// ---- TEST/LOGGING/PROCESSOR/UTILS/FB_LogRecordProcessor_ForBatchInspection.TcPOU
(*
	Processor test double that exposes the batch processor's record queue for assertions.
	Unlike FB_LogRecordProcessor_ForRecordsInspection it does NOT override
	onEmit, so tests exercise the real batch grouping behavior.
*)
FUNCTION_BLOCK FB_LogRecordProcessor_ForBatchInspection EXTENDS FB_LogRecordProcessor_Batch

// explicitly run the batch processor body so tests exercise the flush logic
SUPER^();

PROPERTY records : REFERENCE TO FB_LogRecordQueue
GET
records REF= THIS^._records;
END_GET
END_PROPERTY

END_FUNCTION_BLOCK

// ---- TEST/LOGGING/EXPORTING/FB_TestLogExporters.TcPOU
(* Tests the contract between a caller's batch and a log exporter. *)
FUNCTION_BLOCK FB_TestLogExporters EXTENDS FB_TestSuite

THIS^.testExportSerializesWholeBatch();

(*
	export takes ownership of every record in the caller's batch and passes them to the serializer, so the
	caller holds nothing the exporter will release. Grouping by resource and scope is tested in FB_TestProtoJsonSerializer.
*)
METHOD testExportSerializesWholeBatch : REFERENCE TO FB_Test
VAR CONSTANT
	RECORD_COUNT: UDINT := 2;  // more than one, so the whole batch has to move, not just its head
END_VAR
VAR
	resource: FB_Resource(schemaUrl:='');
	provider: FB_LoggerProvider(resource:=resource);
	scope: FB_InstrumentationScope(name:='exporter.test', version:='1.0.0', schemaUrl:='');
	logger: FB_Logger(scope:=scope, provider:=provider);
	processor: FB_LogRecordProcessor_ForRecordsInspection(
		maxQueueSize:=0,
		scheduledDelayMillis:=1000,
		maxExportBatchSize:=512,
		exporter:=0
	);
	exporter: FB_LogRecordExporter_File_ForSerializationInspection;
	serialized: REFERENCE TO FB_LogRecordProtoJsonSerializer;
	emitSucceeded: BOOL;
	emitFailureReason: E_LoggerFailureReason;
	exporterFailureReason: E_LogRecordExporterFailureReason;
	exportSucceeded: BOOL;
	resourceLogs: SJsonValue;
	_idx: UDINT;
END_VAR
TcUnit.TEST('testExportSerializesWholeBatch');
	// arrange: the processor collects a batch emitted through the logger; its resource and scope do not matter here
	processor.free();
	FOR _idx := 1 TO RECORD_COUNT DO
		emitSucceeded := logger
			.startLogRecord(severityNumber:=E_SeverityNumber.INFO)
			.setTimestamp(TO_ULINT(_idx))
			.emit(failureResult=>emitFailureReason);
		THIS^.AssertTrue(emitSucceeded, 'Expected the logger to emit the record');
	END_FOR
	provider
		.stageProcessor(processor)
		.tick();
	THIS^.AssertEquals_UDINT(RECORD_COUNT, processor.records.count, 'Expected the processor to collect every emitted record');

	// act
	exportSucceeded := processor.exportRecords(exporter:=exporter, failureReason=>exporterFailureReason);

	// assert: the exporter owns the whole batch and serialized it
	THIS^.AssertTrue(
		exportSucceeded
		AND_THEN processor.records.count = 0
		AND_THEN exporterFailureReason = E_LogRecordExporterFailureReason.NA,
		'Expected export to succeed with no failure reason and take every record out of the batch'
	);
	serialized REF= exporter.serializer;
	resourceLogs := serialized.parser.FindMember(serialized.jsonValue, 'resourceLogs');
	THIS^.AssertTrue(resourceLogs <> 0 AND_THEN serialized.parser.IsArray(resourceLogs), 'Expected the exporter to serialize the batch into a resourceLogs array');

	exporter.free();
	processor.free();
TcUnit.TEST_FINISHED();
END_METHOD

END_FUNCTION_BLOCK

// ---- TEST/LOGGING/PROCESSOR/UTILS/FB_LogRecordProcessor_ForRecordsInspection.TcPOU
(* Processor test double that retains emitted records for assertions. *)
// lastOperationSucceeded and failureResult are inherited from FB_LogRecordProcessor_Batch
FUNCTION_BLOCK FB_LogRecordProcessor_ForRecordsInspection EXTENDS FB_LogRecordProcessor_Batch

METHOD exportRecords : BOOL
VAR_INPUT
	exporter: REFERENCE TO FB_LogRecordExporter_Base;
END_VAR
VAR_OUTPUT
	failureReason: E_LogRecordExporterFailureReason;
END_VAR
exportRecords := exporter.export(
	logRecords:=THIS^._records,
	count:=THIS^._records.count,
	failureReason=>failureReason
);
END_METHOD

(*
	Retains every emitted record for assertions, whether or not an exporter is
	bound. FB_LogRecordProcessor_Batch.onEmit deliberately skips the clone and
	the queue push when it has no exporter; this double overrides that so a test
	can collect records and hand them to an exporter itself via exportRecords.
*)
METHOD onEmit
VAR_INPUT
	logRecord: REFERENCE TO FB_LogRecord;
END_VAR
VAR
	_pRecord: POINTER TO FB_LogRecord;
	_cloneFailureResult: E_LogRecordCloneFailureReason;
	_queueFailureReason: E_LogRecordQueueFailureReason;
END_VAR
THIS^.enrich(logRecord);

_pRecord := 0;
IF NOT logRecord.cloneTo(pDest:=_pRecord, failureReason=>_cloneFailureResult) THEN
	IF _pRecord <> 0 THEN _pRecord^.delete(pSelf:=_pRecord); END_IF
	THIS^.lastOperationSucceeded := FALSE;
	THIS^.failureResult := E_LogRecordProcessorFailureReason.RECORD_CLONE_FAILURE;
	RETURN;
END_IF

IF NOT THIS^._records.push(pValue:=_pRecord, failureReason=>_queueFailureReason) THEN
	_pRecord^.delete(pSelf:=_pRecord);
	THIS^.lastOperationSucceeded := FALSE;
	THIS^.failureResult := E_LogRecordProcessorFailureReason.QUEUE_PUSH_FAILURE;
	RETURN;
END_IF

THIS^.lastOperationSucceeded := TRUE;
THIS^.failureResult := E_LogRecordProcessorFailureReason.NA;
END_METHOD

PROPERTY records : REFERENCE TO FB_LogRecordQueue
GET
records REF= THIS^._records;
END_GET
END_PROPERTY

END_FUNCTION_BLOCK

// ---- TEST/LOGGING/EXPORTING/UTILS/FB_LogRecordExporter_File_ForSerializationInspection.TcPOU
(* Exporter test double that serializes accepted records without destination I/O. *)
FUNCTION_BLOCK FB_LogRecordExporter_File_ForSerializationInspection EXTENDS FB_LogRecordExporter_Base
VAR_OUTPUT
	serializer: FB_LogRecordProtoJsonSerializer;
END_VAR
VAR
	_serializationFailureReason: E_ProtoJsonSerializerFailureReason;
END_VAR

METHOD export : BOOL
VAR_IN_OUT
	logRecords: FB_LogRecordQueue;
END_VAR
VAR_INPUT
	count: UDINT;
END_VAR
VAR_OUTPUT
	failureReason: E_LogRecordExporterFailureReason;
END_VAR
_serializationFailureReason := E_ProtoJsonSerializerFailureReason.NA;
export := SUPER^.export(
	logRecords:=logRecords,
	count:=count,
	failureReason=>failureReason
);
IF NOT export THEN
	RETURN;
END_IF

IF NOT THIS^.serializer.serializeLogsData(
	logRecords:=THIS^._records,
	failureReason=>_serializationFailureReason
) THEN
	failureReason := E_LogRecordExporterFailureReason.SERIALIZATION_FAILURE;
	export := FALSE;
END_IF
THIS^.free();
END_METHOD

METHOD isBusy : BOOL
isBusy := FALSE;
END_METHOD

METHOD tick : BOOL
VAR_OUTPUT
	failureReason: E_LogRecordExporterFailureReason;
END_VAR
failureReason := E_LogRecordExporterFailureReason.NA;
tick := TRUE;
END_METHOD

END_FUNCTION_BLOCK

// ---- TEST/LOGGING/LOG_RECORD/FB_TestLogRecord.TcPOU
(* Tests log record ownership and cloning. *)
FUNCTION_BLOCK FB_TestLogRecord EXTENDS FB_TestSuite
VAR_INPUT
END_VAR
VAR_OUTPUT
END_VAR
VAR
END_VAR

THIS^.testCloneToIsIndependent();

(* cloneTo deep copies a record, its resource, scope and every owned value, so a processor can keep the clone after the logger frees the source. Cloning into an assigned destination is refused so the existing record is not leaked. *)
METHOD testCloneToIsIndependent : REFERENCE TO FB_Test
VAR_INPUT
END_VAR
VAR
	resource: FB_Resource('resource.schema');
	provider: FB_LoggerProvider(resource);
	scope: FB_InstrumentationScope('scope.name', '1.0.0', 'scope.schema');
	logger: FB_Logger(scope, provider);
	timestamp: ULINT := 123456789;
	traceIdBytes: ARRAY [0..15] OF BYTE := [0, 1, 2, 3, 4, 5, 6, 7, 8, 9, 10, 11, 12, 13, 14, 15];
	spanIdBytes: ARRAY [0..7] OF BYTE := [16, 17, 18, 19, 20, 21, 22, 23];
	cloneSuccess: BOOL;
	cloneFailureResult: E_LogRecordCloneFailureReason;
	attributesSuccess: BOOL;
	attributesFailureReason: E_AttributesFailureReason;
	pClone: POINTER TO FB_LogRecord;
	pSourceResourceAttribute: POINTER TO FB_KeyValue;
	pClonedResourceAttribute: POINTER TO FB_KeyValue;
	pSourceScopeAttribute: POINTER TO FB_KeyValue;
	pClonedScopeAttribute: POINTER TO FB_KeyValue;
	pSourceRecordAttribute: POINTER TO FB_KeyValue;
	pClonedRecordAttribute: POINTER TO FB_KeyValue;
	pSourceString: POINTER TO FB_String;
	pClonedString: POINTER TO FB_String;
END_VAR
TcUnit.TEST('testCloneToIsIndependent');
	// Arrange: a source record with event name, body, IDs and one attribute at each level
	attributesSuccess := resource.attributes.setStringAttribute(
		key:='resource.key',
		value:='resource.value',
		failureReason=>attributesFailureReason
	);
	THIS^.AssertTrue(attributesSuccess, 'Expected resource attribute creation to succeed');
	attributesSuccess := scope.attributes.setStringAttribute(
		key:='scope.key',
		value:='scope.value',
		failureReason=>attributesFailureReason
	);
	THIS^.AssertTrue(attributesSuccess, 'Expected scope attribute creation to succeed');

	logger
		.startLogRecord(severityNumber:=E_SeverityNumber.INFO)
		.setTimestamp(timestamp)
		.setEventName('record.event')
		.setBody('record.body')
		._setTraceId(ADR(traceIdBytes), SIZEOF(traceIdBytes))
		._setSpanId(ADR(spanIdBytes), SIZEOF(spanIdBytes))
		._setFlags(16#01)  // sampled
		.setStringAttribute('record.key', 'record.value');
	THIS^.AssertTrue(logger.pLogRecord <> 0, 'Expected startLogRecord to build a source log record');

	// Clone: the first clone succeeds, a second into the same destination is refused
	IF logger.pLogRecord <> 0 THEN
		// no builder sets droppedAttributesCount; set by hand so the clone has a non-default value to copy
		logger.pLogRecord^.droppedAttributesCount := 4;
		cloneSuccess := logger.pLogRecord^.cloneTo(
			pDest:=pClone,
			failureReason=>cloneFailureResult
		);
		THIS^.AssertTrue(cloneSuccess, 'Expected log record clone to succeed');
		THIS^.AssertTrue(pClone <> 0, 'Expected a cloned log record');
		THIS^.AssertTrue(pClone <> logger.pLogRecord, 'Expected a distinct log record allocation');

		cloneSuccess := logger.pLogRecord^.cloneTo(
			pDest:=pClone,
			failureReason=>cloneFailureResult
		);
		THIS^.AssertFalse(cloneSuccess, 'Expected cloning into an assigned destination to fail');
		THIS^.AssertTrue(
			cloneFailureResult = E_LogRecordCloneFailureReason.DESTINATION_ALREADY_ASSIGNED,
			'Expected the DESTINATION_ALREADY_ASSIGNED reason when cloning into an assigned destination'
		);
	END_IF

	// Copied fields: equal values, distinct allocations for every owned value
	IF pClone <> 0 AND_THEN logger.pLogRecord <> 0 THEN
		THIS^.AssertTrue(pClone^.severityNumber = logger.pLogRecord^.severityNumber, 'Expected severity number to be cloned');
		THIS^.AssertTrue(pClone^.timestamp = logger.pLogRecord^.timestamp, 'Expected timestamp to be cloned');
		THIS^.AssertEquals_UDINT(logger.pLogRecord^.droppedAttributesCount, pClone^.droppedAttributesCount, 'Expected dropped record attribute count to be cloned');
		THIS^.AssertEquals_STRING(logger.pLogRecord^.resource.schemaUrl, pClone^.resource.schemaUrl, 'Expected resource schema URL to be cloned');
		THIS^.AssertEquals_UDINT(logger.pLogRecord^.resource.droppedAttributesCount, pClone^.resource.droppedAttributesCount, 'Expected dropped resource attribute count to be cloned');
		THIS^.AssertEquals_STRING(logger.pLogRecord^.scope.name, pClone^.scope.name, 'Expected scope name to be cloned');
		THIS^.AssertEquals_STRING(logger.pLogRecord^.scope.version, pClone^.scope.version, 'Expected scope version to be cloned');
		THIS^.AssertEquals_STRING(logger.pLogRecord^.scope.schemaUrl, pClone^.scope.schemaUrl, 'Expected scope schema URL to be cloned');
		THIS^.AssertEquals_UDINT(logger.pLogRecord^.scope.droppedAttributesCount, pClone^.scope.droppedAttributesCount, 'Expected dropped scope attribute count to be cloned');
		THIS^.AssertTrue(pClone^.eventName <> logger.pLogRecord^.eventName, 'Expected event name allocation to be cloned');
		THIS^.AssertTrue(pClone^.eventName^.pString <> logger.pLogRecord^.eventName^.pString, 'Expected event name string allocation to be cloned');
		THIS^.AssertEquals_STRING(logger.pLogRecord^.eventName^.pString^, pClone^.eventName^.pString^, 'Expected event name value to be cloned');
		THIS^.AssertTrue(pClone^.traceId <> logger.pLogRecord^.traceId, 'Expected trace ID allocation to be cloned');
		THIS^.AssertTrue(MEMCMP(ADR(pClone^.traceId^.bytes), ADR(logger.pLogRecord^.traceId^.bytes), SIZEOF(pClone^.traceId^.bytes)) = 0, 'Expected trace ID value to be cloned');
		THIS^.AssertEquals_UDINT(1, pClone^.flags, 'Expected the sampled trace flag to be cloned');
		THIS^.AssertTrue(pClone^.spanId <> logger.pLogRecord^.spanId, 'Expected span ID allocation to be cloned');
		THIS^.AssertTrue(MEMCMP(ADR(pClone^.spanId^.bytes), ADR(logger.pLogRecord^.spanId^.bytes), SIZEOF(pClone^.spanId^.bytes)) = 0, 'Expected span ID value to be cloned');
		THIS^.AssertTrue(pClone^.body <> logger.pLogRecord^.body, 'Expected body allocation to be cloned');
		pSourceString := logger.pLogRecord^.body;
		pClonedString := pClone^.body;
		THIS^.AssertTrue(pClonedString^.pString <> pSourceString^.pString, 'Expected body string allocation to be cloned');
		THIS^.AssertEquals_STRING(pSourceString^.pString^, pClonedString^.pString^, 'Expected body value to be cloned');

		// Attributes: each level's attribute, key and value are new allocations
		logger.pLogRecord^.resource.attributes.reset();
		pClone^.resource.attributes.reset();
		pSourceResourceAttribute := logger.pLogRecord^.resource.attributes.next();
		pClonedResourceAttribute := pClone^.resource.attributes.next();
		THIS^.AssertTrue(pSourceResourceAttribute <> 0, 'Expected the source record to have a resource attribute');
		THIS^.AssertTrue(pClonedResourceAttribute <> 0, 'Expected the cloned record to have a resource attribute');
		IF pSourceResourceAttribute <> 0 AND_THEN pClonedResourceAttribute <> 0 THEN
			THIS^.AssertTrue(pClonedResourceAttribute <> pSourceResourceAttribute, 'Expected resource attribute allocation to be cloned');
			THIS^.AssertTrue(pClonedResourceAttribute^.pKey <> pSourceResourceAttribute^.pKey, 'Expected resource attribute key allocation to be cloned');
			THIS^.AssertTrue(pClonedResourceAttribute^.pVal <> pSourceResourceAttribute^.pVal, 'Expected resource attribute value allocation to be cloned');
		END_IF

		logger.pLogRecord^.scope.attributes.reset();
		pClone^.scope.attributes.reset();
		pSourceScopeAttribute := logger.pLogRecord^.scope.attributes.next();
		pClonedScopeAttribute := pClone^.scope.attributes.next();
		THIS^.AssertTrue(pSourceScopeAttribute <> 0, 'Expected the source record to have a scope attribute');
		THIS^.AssertTrue(pClonedScopeAttribute <> 0, 'Expected the cloned record to have a scope attribute');
		IF pSourceScopeAttribute <> 0 AND_THEN pClonedScopeAttribute <> 0 THEN
			THIS^.AssertTrue(pClonedScopeAttribute <> pSourceScopeAttribute, 'Expected scope attribute allocation to be cloned');
			THIS^.AssertTrue(pClonedScopeAttribute^.pKey <> pSourceScopeAttribute^.pKey, 'Expected scope attribute key allocation to be cloned');
			THIS^.AssertTrue(pClonedScopeAttribute^.pVal <> pSourceScopeAttribute^.pVal, 'Expected scope attribute value allocation to be cloned');
		END_IF

		logger.pLogRecord^.attributes.reset();
		pClone^.attributes.reset();
		pSourceRecordAttribute := logger.pLogRecord^.attributes.next();
		pClonedRecordAttribute := pClone^.attributes.next();
		THIS^.AssertTrue(pSourceRecordAttribute <> 0, 'Expected the source record to have a record attribute');
		THIS^.AssertTrue(pClonedRecordAttribute <> 0, 'Expected the cloned record to have a record attribute');
		IF pSourceRecordAttribute <> 0 AND_THEN pClonedRecordAttribute <> 0 THEN
			THIS^.AssertTrue(pClonedRecordAttribute <> pSourceRecordAttribute, 'Expected record attribute allocation to be cloned');
			THIS^.AssertTrue(pClonedRecordAttribute^.pKey <> pSourceRecordAttribute^.pKey, 'Expected record attribute key allocation to be cloned');
			THIS^.AssertTrue(pClonedRecordAttribute^.pVal <> pSourceRecordAttribute^.pVal, 'Expected record attribute value allocation to be cloned');
		END_IF
	END_IF

	// Independence: the clone keeps its values after the logger frees the source
	logger.free();
	THIS^.AssertTrue(logger.pLogRecord = 0, 'Expected source log record to be deleted');

	IF pClone <> 0 THEN
		THIS^.AssertEquals_STRING('record.event', pClone^.eventName^.pString^, 'Expected cloned event name to survive source deletion');
		pClonedString := pClone^.body;
		THIS^.AssertEquals_STRING('record.body', pClonedString^.pString^, 'Expected cloned body to survive source deletion');
		THIS^.AssertEquals_UDINT(1, pClone^.resource.attributes.count, 'Expected cloned resource attributes to survive source deletion');
		THIS^.AssertEquals_UDINT(1, pClone^.scope.attributes.count, 'Expected cloned scope attributes to survive source deletion');
		THIS^.AssertEquals_UDINT(1, pClone^.attributes.count, 'Expected cloned record attributes to survive source deletion');
		pClone^.delete(pSelf:=pClone);
	END_IF
TcUnit.TEST_FINISHED();
END_METHOD

END_FUNCTION_BLOCK

// ---- TEST/LOGGING/SERIALIZATION/FB_TestProtoJsonSerializer.TcPOU
(* Tests that the base and log-record ProtoJSON serializers write the OTLP/JSON wire form: field encodings, failure reasons, and resource/scope grouping. *)
FUNCTION_BLOCK FB_TestProtoJsonSerializer EXTENDS FB_TestSuite

THIS^.testSerializeNumberValues();
THIS^.testSerializeLogRecord();
THIS^.testSerializeLogRecordWithoutTraceIdOmitsFlags();
THIS^.testSerializeRejectsNullInputs();
THIS^.testSerializeLogsDataGroupsByResourceAndScope();

(* A null log-record pointer or a null member key fails serialization with its own failure reason,
   so a caller can tell a missing record from a serializer misuse instead of writing broken JSON. *)
METHOD testSerializeRejectsNullInputs : REFERENCE TO FB_Test
VAR
	serializer: FB_LogRecordProtoJsonSerializer;
	root: SJsonValue;
	records: SJsonValue;
	pRecord: POINTER TO FB_LogRecord;
	serializationSucceeded: BOOL;
	failureReason: E_ProtoJsonSerializerFailureReason;
END_VAR
TcUnit.TEST('testSerializeRejectsNullInputs');
	root := serializer.parser.NewDocument();
	root := serializer.parser.SetObject(root);
	records := serializer.parser.AddArrayMember(root, 'logRecords', 0);

	// pRecord is deliberately left 0.
	serializationSucceeded := serializer.serializeLogRecord(
		v:=records,
		pLogRecord:=pRecord,
		failureReason=>failureReason
	);
	THIS^.AssertFalse(serializationSucceeded, 'Expected a null log-record pointer to fail serialization');
	THIS^.AssertTrue(
		failureReason = E_ProtoJsonSerializerFailureReason.LOG_RECORD_POINTER_NULL,
		'Expected LOG_RECORD_POINTER_NULL as the failure reason for a null log record'
	);

	// pKey is deliberately 0.
	serializationSucceeded := serializer.serializeUint32Value(
		v:=root,
		pKey:=0,
		val:=1,
		failureReason=>failureReason
	);
	THIS^.AssertFalse(serializationSucceeded, 'Expected a null JSON member key to fail serialization');
	THIS^.AssertTrue(
		failureReason = E_ProtoJsonSerializerFailureReason.KEY_POINTER_NULL,
		'Expected KEY_POINTER_NULL as the failure reason for a null member key'
	);
TcUnit.TEST_FINISHED();
END_METHOD

(* A record built through the logger serializes every field in its OTLP/JSON form: enums and fixed32 as numbers,
   64-bit integers as decimal strings, trace and span IDs as hex, and values as typed AnyValue objects. *)
METHOD testSerializeLogRecord : REFERENCE TO FB_Test
VAR
	resource: FB_Resource(schemaUrl:='');
	provider: FB_LoggerProvider(resource:=resource);
	scope: FB_InstrumentationScope(name:='motor1', version:='0.0.1a', schemaUrl:='');
	logger: FB_Logger(scope:=scope, provider:=provider);
	processor: FB_LogRecordProcessor_ForRecordInspection(0);
	serializer: FB_LogRecordProtoJsonSerializer();
	emitSuccess: BOOL;
	emitFailureResult: E_LoggerFailureReason;
	timestamp: ULINT := 1581452773000000789;
	traceId: ARRAY [0..15] OF BYTE := [0, 1, 2, 3, 4, 5, 6, 7, 8, 9, 10, 11, 12, 13, 14, 15];
	spanId: ARRAY [0..7] OF BYTE := [16, 17, 18, 19, 20, 21, 22, 23];
	durationMs: DINT := 42;
	temperature: LREAL := 21.5;
	pRecord: POINTER TO FB_LogRecord;
	root: SJsonValue;
	records: SJsonValue;
	obj: SJsonValue;
	member: SJsonValue;
	attributes: SJsonValue;
	attribute: SJsonValue;
	value: SJsonValue;
	actualString: STRING;
	serializationSucceeded: BOOL;
	serializerFailureReason: E_ProtoJsonSerializerFailureReason;
END_VAR
TcUnit.TEST('testSerializeLogRecord');
	processor.free();
	logger.free();

	// Create a representative record through the public logger API.
	logger
		.startLogRecord(severityNumber:=E_SeverityNumber.DEBUG)
		.setTimestamp(timestamp)
		.setEventName('Serialization Event')
		.setBody('This is a body string value')
		._setTraceId(ADR(traceId), SIZEOF(traceId))
		._setSpanId(ADR(spanId), SIZEOF(spanId))
		._setFlags(16#01)  // sampled
		.setStringAttribute('stats.label', 'pVal')
		.setNumberAttribute('stats.duration_ms', durationMs)
		.setNumberAttribute('stats.temperature', temperature);
	THIS^.AssertTrue(logger.pLogRecord <> 0, 'Expected the logger to hold a log record before emission');
	IF logger.pLogRecord <> 0 THEN
		// no builder sets droppedAttributesCount; set by hand to check it is written
		logger.pLogRecord^.droppedAttributesCount := 2;
	END_IF

	emitSuccess := logger.emit(failureResult=>emitFailureResult);
	THIS^.AssertTrue(emitSuccess, 'Expected log record emission to succeed');
	provider
		.stageProcessor(processor)
		.tick();
	THIS^.AssertTrue(processor.lastOperationSucceeded, 'Expected the inspection processor to capture the emitted record');
	THIS^.AssertTrue(logger.pLogRecord = 0, 'Expected emit to release the logger-owned record');
	pRecord := processor.pop();
	THIS^.AssertTrue(pRecord <> 0, 'Expected the processor to return the emitted record');
	IF pRecord <> 0 THEN

	// serializeLogRecord appends one LogRecord object to the supplied JSON array.
	root := serializer.parser.NewDocument();
	serializer.parser.SetObject(root);
	records := serializer.parser.AddArrayMember(root, 'logRecords', 0);
	serializationSucceeded := serializer.serializeLogRecord(
		v:=records,
		pLogRecord:=pRecord,
		failureReason=>serializerFailureReason
	);
	THIS^.AssertTrue(
		serializationSucceeded AND_THEN serializerFailureReason = E_ProtoJsonSerializerFailureReason.NA,
		'Expected LogRecord serialization to succeed without a failure reason'
	);
	obj := serializer.parser.GetArrayValueByIdx(records, 0);
		THIS^.AssertTrue(serializer.parser.IsObject(obj), 'Expected the logRecords array to hold one LogRecord object');

		// OTLP/JSON encodes enums and fixed32 values as numbers.
		// 5 is DEBUG; flags 1 is the sampled trace flag of the record's span.
		member := serializer.parser.FindMember(obj, 'severityNumber');
		THIS^.AssertEquals_UDINT(5, serializer.parser.GetUint(member), 'Expected severityNumber 5 (DEBUG) as a JSON number');
		actualString := serializer.parser.GetString(serializer.parser.FindMember(obj, 'severityText'));
		THIS^.AssertEquals_STRING('DEBUG', actualString, 'Expected severityText to be the severity enum name');
		THIS^.AssertEquals_UDINT(1, serializer.parser.GetUint(serializer.parser.FindMember(obj, 'flags')), 'Expected flags 1 (sampled) as a JSON number');
		THIS^.AssertEquals_UDINT(2, serializer.parser.GetUint(serializer.parser.FindMember(obj, 'droppedAttributesCount')), 'Expected droppedAttributesCount 2 as a JSON number');

		// OTLP/JSON encodes 64-bit integers as decimal strings and trace/span IDs as hex.
		actualString := serializer.parser.GetString(serializer.parser.FindMember(obj, 'timeUnixNano'));
		THIS^.AssertEquals_STRING('1581452773000000789', actualString, 'Expected string-encoded timeUnixNano');
		actualString := serializer.parser.GetString(serializer.parser.FindMember(obj, 'traceId'));
		THIS^.AssertEquals_STRING('000102030405060708090A0B0C0D0E0F', actualString, 'Expected hex-encoded traceId');
		actualString := serializer.parser.GetString(serializer.parser.FindMember(obj, 'spanId'));
		THIS^.AssertEquals_STRING('1011121314151617', actualString, 'Expected hex-encoded spanId');

		// Event name and body.
		actualString := serializer.parser.GetString(serializer.parser.FindMember(obj, 'eventName'));
		THIS^.AssertEquals_STRING('Serialization Event', actualString, 'Expected eventName to be written as set');
		value := serializer.parser.FindMember(serializer.parser.FindMember(obj, 'body'), 'stringValue');
		actualString := serializer.parser.GetString(value);
		THIS^.AssertEquals_STRING('This is a body string value', actualString, 'Expected AnyValue string body');

		// Attributes keep insertion order; each value is a typed AnyValue, with intValue as a decimal string.
		attributes := serializer.parser.FindMember(obj, 'attributes');
		THIS^.AssertTrue(serializer.parser.IsArray(attributes), 'Expected attributes to be a JSON array');
		attribute := serializer.parser.GetArrayValueByIdx(attributes, 0);
		actualString := serializer.parser.GetString(serializer.parser.FindMember(attribute, 'key'));
		THIS^.AssertEquals_STRING('stats.label', actualString, 'Expected string attribute key');
		value := serializer.parser.FindMember(serializer.parser.FindMember(attribute, 'value'), 'stringValue');
		actualString := serializer.parser.GetString(value);
		THIS^.AssertEquals_STRING('pVal', actualString, 'Expected string attribute AnyValue');
		attribute := serializer.parser.GetArrayValueByIdx(attributes, 1);
		actualString := serializer.parser.GetString(serializer.parser.FindMember(attribute, 'key'));
		THIS^.AssertEquals_STRING('stats.duration_ms', actualString, 'Expected numeric attribute key');
		value := serializer.parser.FindMember(serializer.parser.FindMember(attribute, 'value'), 'intValue');
		actualString := serializer.parser.GetString(value);
		THIS^.AssertEquals_STRING('42', actualString, 'Expected numeric attribute AnyValue');
		attribute := serializer.parser.GetArrayValueByIdx(attributes, 2);
		actualString := serializer.parser.GetString(serializer.parser.FindMember(attribute, 'key'));
		THIS^.AssertEquals_STRING('stats.temperature', actualString, 'Expected floating attribute key');
		value := serializer.parser.FindMember(serializer.parser.FindMember(attribute, 'value'), 'doubleValue');
		THIS^.AssertTrue(serializer.parser.IsDouble(value) AND_THEN serializer.parser.GetDouble(value) = 21.5, 'Expected floating attribute AnyValue');
	END_IF

	IF pRecord <> 0 THEN pRecord^.delete(pSelf:=pRecord); END_IF
	processor.free();
	logger.free();

TcUnit.TEST_FINISHED();
END_METHOD

(* A record without a trace id belongs to no trace, so the serializer leaves out flags even when the record holds some,
   along with traceId and spanId. The record stores flags as set; omitting them is the serializer's decision. *)
METHOD testSerializeLogRecordWithoutTraceIdOmitsFlags : REFERENCE TO FB_Test
VAR
	resource: FB_Resource(schemaUrl:='');
	provider: FB_LoggerProvider(resource:=resource);
	scope: FB_InstrumentationScope(name:='motor1', version:='0.0.1a', schemaUrl:='');
	logger: FB_Logger(scope:=scope, provider:=provider);
	processor: FB_LogRecordProcessor_ForRecordInspection(0);
	serializer: FB_LogRecordProtoJsonSerializer();
	emitSuccess: BOOL;
	emitFailureResult: E_LoggerFailureReason;
	pRecord: POINTER TO FB_LogRecord;
	root: SJsonValue;
	records: SJsonValue;
	obj: SJsonValue;
	serializationSucceeded: BOOL;
	serializerFailureReason: E_ProtoJsonSerializerFailureReason;
END_VAR
TcUnit.TEST('testSerializeLogRecordWithoutTraceIdOmitsFlags');
	emitSuccess := logger
		.startLogRecord(severityNumber:=E_SeverityNumber.INFO)
		._setFlags(16#01)  // sampled, but no trace id
		.emit(failureResult=>emitFailureResult);
	THIS^.AssertTrue(emitSuccess, 'Expected log record emission to succeed');
	provider
		.stageProcessor(processor)
		.tick();
	pRecord := processor.pop();
	THIS^.AssertTrue(pRecord <> 0, 'Expected the processor to return the emitted record');
	IF pRecord <> 0 THEN
		THIS^.AssertEquals_UDINT(1, pRecord^.flags, 'Expected the record to keep the flags it was given');

		root := serializer.parser.NewDocument();
		serializer.parser.SetObject(root);
		records := serializer.parser.AddArrayMember(root, 'logRecords', 0);
		serializationSucceeded := serializer.serializeLogRecord(
			v:=records,
			pLogRecord:=pRecord,
			failureReason=>serializerFailureReason
		);
		THIS^.AssertTrue(serializationSucceeded, 'Expected LogRecord serialization to succeed');
		obj := serializer.parser.GetArrayValueByIdx(records, 0);
		THIS^.AssertTrue(serializer.parser.IsObject(obj), 'Expected the logRecords array to hold one LogRecord object');
		THIS^.AssertTrue(serializer.parser.FindMember(obj, 'flags') = 0, 'Expected no flags member without a trace id');
		THIS^.AssertTrue(serializer.parser.FindMember(obj, 'traceId') = 0, 'Expected no traceId member');
		THIS^.AssertTrue(serializer.parser.FindMember(obj, 'spanId') = 0, 'Expected no spanId member');
		pRecord^.delete(pSelf:=pRecord);
	END_IF
	processor.free();
TcUnit.TEST_FINISHED();
END_METHOD

(* serializeLogsData groups interleaved records into one ResourceLogs per resource and one ScopeLogs per scope,
   in first-seen order with records kept in arrival order, and drains the queue it is given. *)
METHOD testSerializeLogsDataGroupsByResourceAndScope : REFERENCE TO FB_Test
VAR
	resourceB: FB_Resource('resource.b');
	resourceA: FB_Resource('resource.a');
	resourceC: FB_Resource('resource.c');
	providerB: FB_LoggerProvider(resource:=resourceB);
	providerA: FB_LoggerProvider(resource:=resourceA);
	providerC: FB_LoggerProvider(resource:=resourceC);
	scopeB: FB_InstrumentationScope('scope.b', '1.0.0', 'scope.b.schema');
	scopeA: FB_InstrumentationScope('scope.a', '1.0.0', 'scope.a.schema');
	scopeC: FB_InstrumentationScope('scope.c', '1.0.0', 'scope.c.schema');
	loggerBb: FB_Logger(scope:=scopeB, provider:=providerB);
	loggerBa: FB_Logger(scope:=scopeA, provider:=providerB);
	loggerAc: FB_Logger(scope:=scopeC, provider:=providerA);
	loggerAb: FB_Logger(scope:=scopeB, provider:=providerA);
	loggerCa: FB_Logger(scope:=scopeA, provider:=providerC);
	processor: FB_LogRecordProcessor_ForRecordsInspection(
		maxQueueSize:=0,
		scheduledDelayMillis:=1000,
		maxExportBatchSize:=512,
		exporter:=0
	);
	queue: REFERENCE TO FB_LogRecordQueue;
	serializer: FB_LogRecordProtoJsonSerializer;
	emitSucceeded: BOOL;
	_idx: UDINT;
	resourceLogs: SJsonValue;
	resourceObj: SJsonValue;
	scopeLogs: SJsonValue;
	scopeObj: SJsonValue;
	logRecords: SJsonValue;
	recordObj: SJsonValue;
	actualString: STRING;
	serializationSucceeded: BOOL;
	serializerFailureReason: E_ProtoJsonSerializerFailureReason;
END_VAR
TcUnit.TEST('testSerializeLogsDataGroupsByResourceAndScope');
	processor.free();
	queue REF= processor.records;

	// ---- Arrange: eight records with interleaved resource/scope pairs ----
	// Each logger is one resource/scope pair, named resource then scope (loggerBa is resource B, scope A).
	// The timestamp is the record number, so each record can be identified in the output.
	//   record:   1  2  3  4  5  6  7  8
	//   resource: B  A  C  B  C  A  B  A
	//   scope:    B  C  A  A  A  B  B  C
	FOR _idx := 1 TO 8 DO
		CASE _idx OF
			1, 7: emitSucceeded := THIS^._emitRecord(logger:=loggerBb, provider:=providerB, processor:=processor, timestamp:=_idx);
			4:    emitSucceeded := THIS^._emitRecord(logger:=loggerBa, provider:=providerB, processor:=processor, timestamp:=_idx);
			2, 8: emitSucceeded := THIS^._emitRecord(logger:=loggerAc, provider:=providerA, processor:=processor, timestamp:=_idx);
			6:    emitSucceeded := THIS^._emitRecord(logger:=loggerAb, provider:=providerA, processor:=processor, timestamp:=_idx);
			3, 5: emitSucceeded := THIS^._emitRecord(logger:=loggerCa, provider:=providerC, processor:=processor, timestamp:=_idx);
		END_CASE
		THIS^.AssertTrue(emitSucceeded, CONCAT('Expected record ', CONCAT(UDINT_TO_STRING(_idx), ' to reach the processor')));
	END_FOR
	THIS^.AssertEquals_UDINT(8, queue.count, 'Expected eight records queued before serialization');

	// ---- Act ----
	serializationSucceeded := serializer.serializeLogsData(
		logRecords:=queue,
		failureReason=>serializerFailureReason
	);
	THIS^.AssertTrue(
		serializationSucceeded AND_THEN serializerFailureReason = E_ProtoJsonSerializerFailureReason.NA,
		'Expected LogsData serialization to succeed without a failure reason'
	);
	THIS^.AssertEquals_UDINT(0, queue.count, 'Expected the serializer to drain the queue it was given');

	// ---- Assert: three ResourceLogs groups in first-seen order B, A, C ----
	resourceLogs := serializer.parser.FindMember(serializer.jsonValue, 'resourceLogs');
	THIS^.AssertTrue(resourceLogs <> 0 AND_THEN serializer.parser.IsArray(resourceLogs), 'Expected resourceLogs to be a JSON array');

	THIS^.AssertTrue(serializer.parser.GetArrayValueByIdx(resourceLogs, 3) = 0, 'Expected exactly three ResourceLogs groups');

	// Resource B was seen first. Its scope B records remain in arrival order,
	// followed by the later first-seen scope A group.
	resourceObj := serializer.parser.GetArrayValueByIdx(resourceLogs, 0);
	actualString := serializer.parser.GetString(serializer.parser.FindMember(resourceObj, 'schemaUrl'));
	THIS^.AssertEquals_STRING('resource.b', actualString, 'Expected resource B as the first ResourceLogs group');
	scopeLogs := serializer.parser.FindMember(resourceObj, 'scopeLogs');
	scopeObj := serializer.parser.GetArrayValueByIdx(scopeLogs, 0);

	actualString := serializer.parser.GetString(serializer.parser.FindMember(serializer.parser.FindMember(scopeObj, 'scope'), 'name'));
	THIS^.AssertEquals_STRING('scope.b', actualString, 'Expected scope B as the first scope of resource B');
	logRecords := serializer.parser.FindMember(scopeObj, 'logRecords');
	recordObj := serializer.parser.GetArrayValueByIdx(logRecords, 0);

	actualString := serializer.parser.GetString(serializer.parser.FindMember(recordObj, 'timeUnixNano'));
	THIS^.AssertEquals_STRING('1', actualString, 'Expected record 1 first in resource B scope B');
	recordObj := serializer.parser.GetArrayValueByIdx(logRecords, 1);
	actualString := serializer.parser.GetString(serializer.parser.FindMember(recordObj, 'timeUnixNano'));
	THIS^.AssertEquals_STRING('7', actualString, 'Expected record 7 second in resource B scope B');
	THIS^.AssertTrue(serializer.parser.GetArrayValueByIdx(logRecords, 2) = 0, 'Expected exactly two records in resource B scope B');

	scopeObj := serializer.parser.GetArrayValueByIdx(scopeLogs, 1);
	actualString := serializer.parser.GetString(serializer.parser.FindMember(serializer.parser.FindMember(scopeObj, 'scope'), 'name'));
	THIS^.AssertEquals_STRING('scope.a', actualString, 'Expected scope A as the second scope of resource B');
	logRecords := serializer.parser.FindMember(scopeObj, 'logRecords');
	recordObj := serializer.parser.GetArrayValueByIdx(logRecords, 0);

	actualString := serializer.parser.GetString(serializer.parser.FindMember(recordObj, 'timeUnixNano'));
	THIS^.AssertEquals_STRING('4', actualString, 'Expected record 4 in resource B scope A');
	THIS^.AssertTrue(serializer.parser.GetArrayValueByIdx(logRecords, 1) = 0, 'Expected exactly one record in resource B scope A');
	THIS^.AssertTrue(serializer.parser.GetArrayValueByIdx(scopeLogs, 2) = 0, 'Expected exactly two scopes for resource B');

	// Resource A was seen second. Its repeated scope C records are one group.
	resourceObj := serializer.parser.GetArrayValueByIdx(resourceLogs, 1);
	actualString := serializer.parser.GetString(serializer.parser.FindMember(resourceObj, 'schemaUrl'));
	THIS^.AssertEquals_STRING('resource.a', actualString, 'Expected resource A as the second ResourceLogs group');
	scopeLogs := serializer.parser.FindMember(resourceObj, 'scopeLogs');
	scopeObj := serializer.parser.GetArrayValueByIdx(scopeLogs, 0);

	actualString := serializer.parser.GetString(serializer.parser.FindMember(serializer.parser.FindMember(scopeObj, 'scope'), 'name'));
	THIS^.AssertEquals_STRING('scope.c', actualString, 'Expected scope C as the first scope of resource A');
	logRecords := serializer.parser.FindMember(scopeObj, 'logRecords');
	recordObj := serializer.parser.GetArrayValueByIdx(logRecords, 0);

	actualString := serializer.parser.GetString(serializer.parser.FindMember(recordObj, 'timeUnixNano'));
	THIS^.AssertEquals_STRING('2', actualString, 'Expected record 2 first in resource A scope C');
	recordObj := serializer.parser.GetArrayValueByIdx(logRecords, 1);

	actualString := serializer.parser.GetString(serializer.parser.FindMember(recordObj, 'timeUnixNano'));
	THIS^.AssertEquals_STRING('8', actualString, 'Expected record 8 second in resource A scope C');
	THIS^.AssertTrue(serializer.parser.GetArrayValueByIdx(logRecords, 2) = 0, 'Expected exactly two records in resource A scope C');

	scopeObj := serializer.parser.GetArrayValueByIdx(scopeLogs, 1);
	actualString := serializer.parser.GetString(serializer.parser.FindMember(serializer.parser.FindMember(scopeObj, 'scope'), 'name'));
	THIS^.AssertEquals_STRING('scope.b', actualString, 'Expected scope B as the second scope of resource A');
	logRecords := serializer.parser.FindMember(scopeObj, 'logRecords');
	recordObj := serializer.parser.GetArrayValueByIdx(logRecords, 0);
	actualString := serializer.parser.GetString(serializer.parser.FindMember(recordObj, 'timeUnixNano'));
	THIS^.AssertEquals_STRING('6', actualString, 'Expected record 6 in resource A scope B');
	THIS^.AssertTrue(serializer.parser.GetArrayValueByIdx(logRecords, 1) = 0, 'Expected exactly one record in resource A scope B');
	THIS^.AssertTrue(serializer.parser.GetArrayValueByIdx(scopeLogs, 2) = 0, 'Expected exactly two scopes for resource A');

	// Resource C was seen third and its non-adjacent records share one scope.
	resourceObj := serializer.parser.GetArrayValueByIdx(resourceLogs, 2);
	actualString := serializer.parser.GetString(serializer.parser.FindMember(resourceObj, 'schemaUrl'));
	THIS^.AssertEquals_STRING('resource.c', actualString, 'Expected resource C as the third ResourceLogs group');
	scopeLogs := serializer.parser.FindMember(resourceObj, 'scopeLogs');
	scopeObj := serializer.parser.GetArrayValueByIdx(scopeLogs, 0);
	actualString := serializer.parser.GetString(serializer.parser.FindMember(serializer.parser.FindMember(scopeObj, 'scope'), 'name'));
	THIS^.AssertEquals_STRING('scope.a', actualString, 'Expected scope A as the only scope of resource C');
	logRecords := serializer.parser.FindMember(scopeObj, 'logRecords');
	recordObj := serializer.parser.GetArrayValueByIdx(logRecords, 0);
	actualString := serializer.parser.GetString(serializer.parser.FindMember(recordObj, 'timeUnixNano'));
	THIS^.AssertEquals_STRING('3', actualString, 'Expected record 3 first in resource C scope A');
	recordObj := serializer.parser.GetArrayValueByIdx(logRecords, 1);
	actualString := serializer.parser.GetString(serializer.parser.FindMember(recordObj, 'timeUnixNano'));
	THIS^.AssertEquals_STRING('5', actualString, 'Expected record 5 second in resource C scope A');
	THIS^.AssertTrue(serializer.parser.GetArrayValueByIdx(logRecords, 2) = 0, 'Expected exactly two records in resource C scope A');
	THIS^.AssertTrue(serializer.parser.GetArrayValueByIdx(scopeLogs, 1) = 0, 'Expected exactly one scope for resource C');

	processor.free();
TcUnit.TEST_FINISHED();
END_METHOD

(* Integers up to 32 bits and finite floats are written as JSON numbers, while 64-bit integers and
   NaN/Infinity are written as strings, as ProtoJSON requires so that no value loses precision or breaks JSON. *)
METHOD testSerializeNumberValues : REFERENCE TO FB_Test
VAR
	serializer: FB_BaseProtoJsonSerializer;
	root: SJsonValue;
	nSInt: SINT := -12;
	nInt: INT := -1234;
	nDInt: DINT := -123456789;
	nLInt: LINT := -9007199254740993; // -(2^53 + 1): cannot be held exactly by a JSON (double) number
	nUSInt: USINT := 12;
	nUInt: UINT := 1234;
	nUDInt: UDINT := 4000000000;
	nULInt: ULINT := 18000000000000000000; // above 2^63, so it only fits an unsigned 64-bit integer
	fReal: REAL := 42.25;
	fLReal: LREAL := -24.5;
	fNaN: LREAL;
	fPositiveInfinity: LREAL;
	fNegativeInfinity: LREAL;
	// IEEE 754 double bit patterns; ST has no literals for these values.
	nNaNBits: LWORD := LWORD#16#7FF8000000000000;
	nPositiveInfinityBits: LWORD := LWORD#16#7FF0000000000000;
	nNegativeInfinityBits: LWORD := LWORD#16#FFF0000000000000;
	member: SJsonValue;
	actualString: STRING;
END_VAR
TcUnit.TEST('testSerializeNumberValues');
	root := serializer.parser.NewDocument();
	serializer.parser.SetObject(root);

	// serializeNumberValue takes ANY_NUM and dispatches on the actual type.
	THIS^.AssertTrue(serializer.serializeNumberValue(root, ADR('sintValue'), nSInt), 'Expected a SINT to serialize');
	THIS^.AssertTrue(serializer.serializeNumberValue(root, ADR('intValue'), nInt), 'Expected an INT to serialize');
	THIS^.AssertTrue(serializer.serializeNumberValue(root, ADR('dintValue'), nDInt), 'Expected a DINT to serialize');
	THIS^.AssertTrue(serializer.serializeNumberValue(root, ADR('lintValue'), nLInt), 'Expected a LINT to serialize');
	THIS^.AssertTrue(serializer.serializeNumberValue(root, ADR('usintValue'), nUSInt), 'Expected a USINT to serialize');
	THIS^.AssertTrue(serializer.serializeNumberValue(root, ADR('uintValue'), nUInt), 'Expected a UINT to serialize');
	THIS^.AssertTrue(serializer.serializeNumberValue(root, ADR('udintValue'), nUDInt), 'Expected a UDINT to serialize');
	THIS^.AssertTrue(serializer.serializeNumberValue(root, ADR('ulintValue'), nULInt), 'Expected a ULINT to serialize');
	THIS^.AssertTrue(serializer.serializeNumberValue(root, ADR('realValue'), fReal), 'Expected a REAL to serialize');
	THIS^.AssertTrue(serializer.serializeNumberValue(root, ADR('lrealValue'), fLReal), 'Expected an LREAL to serialize');

	THIS^.AssertEquals_DINT(-12, serializer.parser.GetInt(serializer.parser.FindMember(root, 'sintValue')), 'Expected SINT as a JSON number');
	THIS^.AssertEquals_DINT(-1234, serializer.parser.GetInt(serializer.parser.FindMember(root, 'intValue')), 'Expected INT as a JSON number');
	THIS^.AssertEquals_DINT(-123456789, serializer.parser.GetInt(serializer.parser.FindMember(root, 'dintValue')), 'Expected DINT as a JSON number');
	actualString := serializer.parser.GetString(serializer.parser.FindMember(root, 'lintValue'));
	THIS^.AssertEquals_STRING('-9007199254740993', actualString, 'Expected LINT as a decimal JSON string');
	THIS^.AssertEquals_UDINT(12, serializer.parser.GetUint(serializer.parser.FindMember(root, 'usintValue')), 'Expected USINT as a JSON number');
	THIS^.AssertEquals_UDINT(1234, serializer.parser.GetUint(serializer.parser.FindMember(root, 'uintValue')), 'Expected UINT as a JSON number');
	THIS^.AssertEquals_UDINT(4000000000, serializer.parser.GetUint(serializer.parser.FindMember(root, 'udintValue')), 'Expected UDINT as a JSON number');
	actualString := serializer.parser.GetString(serializer.parser.FindMember(root, 'ulintValue'));
	THIS^.AssertEquals_STRING('18000000000000000000', actualString, 'Expected ULINT as a decimal JSON string');
	member := serializer.parser.FindMember(root, 'realValue');
	THIS^.AssertTrue(serializer.parser.IsDouble(member) AND_THEN serializer.parser.GetDouble(member) = 42.25, 'Expected REAL as a JSON number');
	member := serializer.parser.FindMember(root, 'lrealValue');
	THIS^.AssertTrue(serializer.parser.IsDouble(member) AND_THEN serializer.parser.GetDouble(member) = -24.5, 'Expected LREAL as a JSON number');

	// ProtoJSON requires special floating-point values to be quoted strings.
	MEMCPY(ADR(fNaN), ADR(nNaNBits), SIZEOF(fNaN));
	MEMCPY(ADR(fPositiveInfinity), ADR(nPositiveInfinityBits), SIZEOF(fPositiveInfinity));
	MEMCPY(ADR(fNegativeInfinity), ADR(nNegativeInfinityBits), SIZEOF(fNegativeInfinity));
	serializer.serializeNumberValue(root, ADR('nanValue'), fNaN);
	serializer.serializeNumberValue(root, ADR('positiveInfinityValue'), fPositiveInfinity);
	serializer.serializeNumberValue(root, ADR('negativeInfinityValue'), fNegativeInfinity);
	actualString := serializer.parser.GetString(serializer.parser.FindMember(root, 'nanValue'));
	THIS^.AssertEquals_STRING('NaN', actualString, 'Expected NaN as the quoted string NaN');
	actualString := serializer.parser.GetString(serializer.parser.FindMember(root, 'positiveInfinityValue'));
	THIS^.AssertEquals_STRING('Infinity', actualString, 'Expected positive infinity as the quoted string Infinity');
	actualString := serializer.parser.GetString(serializer.parser.FindMember(root, 'negativeInfinityValue'));
	THIS^.AssertEquals_STRING('-Infinity', actualString, 'Expected negative infinity as the quoted string -Infinity');

TcUnit.TEST_FINISHED();
END_METHOD

(*
	Emits one INFO record stamped with timestamp through logger, then ticks its provider with the
	processor staged, so the record reaches the processor now and records keep their emit order
	across providers.
*)
METHOD _emitRecord : BOOL
VAR_INPUT
	logger: REFERENCE TO FB_Logger;
	provider: REFERENCE TO FB_LoggerProvider;
	processor: REFERENCE TO FB_LogRecordProcessor_Base;
	timestamp: ULINT;
END_VAR
VAR
	emitFailureReason: E_LoggerFailureReason;
END_VAR
_emitRecord := logger
	.startLogRecord(severityNumber:=E_SeverityNumber.INFO)
	.setTimestamp(timestamp)
	.emit(failureResult=>emitFailureReason);
_emitRecord := _emitRecord AND_THEN provider
	.stageProcessor(processor)
	.tick();
END_METHOD

END_FUNCTION_BLOCK

// ---- TEST/LOGGING/PROCESSOR/UTILS/FB_LogRecordProcessor_ForRecordInspection.TcPOU
(* Processor test double that retains one emitted record for assertions. *)
FUNCTION_BLOCK FB_LogRecordProcessor_ForRecordInspection EXTENDS FB_LogRecordProcessor_Simple
VAR_OUTPUT
	record: POINTER TO FB_LogRecord;
	lastOperationSucceeded: BOOL := FALSE;
	failureResult: E_LogRecordCloneFailureReason;
END_VAR

METHOD free
IF THIS^.record <> 0 THEN
	THIS^.record^.delete(pSelf:=THIS^.record);
END_IF
END_METHOD

METHOD onEmit
VAR_INPUT
	logRecord: REFERENCE TO FB_LogRecord;
END_VAR
THIS^.free();
THIS^.lastOperationSucceeded := logRecord.cloneTo(
	pDest:=THIS^.record,
	failureReason=>THIS^.failureResult
);
END_METHOD

METHOD pop : POINTER TO FB_LogRecord
pop := THIS^.record;
THIS^.record := 0;
END_METHOD

END_FUNCTION_BLOCK

// ---- TEST/LOGGING/EXPORTING/FB_TestFileExporter.TcPOU
(* Tests that the file log exporter writes processed batches to disk. *)
FUNCTION_BLOCK FB_TestFileExporter EXTENDS FB_TestSuite
VAR
	_resource:		FB_Resource(schemaUrl:='');
	_exporter: 		FB_LogRecordExporter_File(filepath:='C:\Users\samue\Desktop\programming projects\TcOtlp\logs.jsonl');
	_processor:		FB_LogRecordProcessor_ForRecordsInspection(
		maxQueueSize:=0,
		scheduledDelayMillis:=1000,
		maxExportBatchSize:=512,
		exporter:=0
	);
	_provider:		FB_LoggerProvider(resource:=_resource);
	_scope1:			FB_InstrumentationScope(name:='scope1', version:='0.0.1', schemaUrl:='');
	_logger1:		FB_Logger(scope:=_scope1, provider:=_provider);
	_scope2:			FB_InstrumentationScope(name:='scope2', version:='0.0.1', schemaUrl:='');
	_logger2:		FB_Logger(scope:=_scope2, provider:=_provider);
END_VAR

THIS^.testExportBatchedLogRecords(cleanup:=FALSE);

(*
	Records emitted through two loggers reach the file as one batch, and a batch handed over in the
	scan the previous one finished still starts, so back-to-back flushes never stall the file exporter.
*)
METHOD testExportBatchedLogRecords : REFERENCE TO FB_Test

VAR_INPUT
	cleanup: BOOL := TRUE;  // FALSE keeps logs.jsonl on disk for manual inspection
END_VAR

VAR CONSTANT
	_filepath: STRING := 'C:\Users\samue\Desktop\programming projects\TcOtlp\logs.jsonl';
	MAX_CYCLES: UDINT := 1000;
END_VAR

VAR_INST
	_cycles: 		UDINT;
	_state:			USINT;
	_redelivered:	BOOL;  // a second batch was exported in the scan the first finished
	_fileFinder: 	FB_EnumFindFileEntry;
	_fileDeleter:	FB_FileDelete;
END_VAR

VAR
	_num: UINT;
	_fileSize: ULINT;
	_exportSucceeded: BOOL;
	_exportCallSucceeded: BOOL;
	_firstEmitSucceeded: BOOL;
	_secondEmitSucceeded: BOOL;
	_thirdEmitSucceeded: BOOL;
	_loggerFailureResult: E_LoggerFailureReason;
	_exporterFailureReason: E_LogRecordExporterFailureReason;
	_timestamp: ULINT := ULINT#1581452773000000789;
	_traceId: ARRAY[0..ValueFactory.nTraceIdBytes-1] OF BYTE := [0, 1, 2, 3, 4, 5, 6, 7, 8, 9, 10, 11, 12, 13, 14, 15];
	_spanId: ARRAY[0..ValueFactory.nSpanIdBytes-1] OF BYTE := [16, 17, 18, 19, 20, 21, 22, 23];
END_VAR
TcUnit.TEST('testExportBatchedLogRecords');
	CASE _state OF
		0: // emit three records through two loggers; the processor captures them without exporting
			_cycles := 0;
			_redelivered := FALSE;
			_processor.free();
			_logger1.free();
			// _resource persists across test re-runs; only add the attribute once
			IF _resource.attributes.count = 0 THEN
				_resource.attributes.setStringAttribute('host.id', 'PLC1');
			END_IF
			_num := 1;
			_firstEmitSucceeded := _logger1
				.startLogRecord(severityNumber:=E_SeverityNumber.DEBUG)
				.setTimestamp(_timestamp)
				.setBody('First batched log record')
				.setEventName('BatchRecord1')
				._setTraceId(ADR(_traceId), SIZEOF(_traceId))
				._setSpanId(ADR(_spanId), SIZEOF(_spanId))
				.setStringAttribute('batch.position', 'first')
				.setNumberAttribute('batch.positionNum', _num)
				.emit(failureResult=>_loggerFailureResult);
			_num := 2;
			_secondEmitSucceeded := _logger2
				.startLogRecord(severityNumber:=E_SeverityNumber.INFO)
				.setTimestamp(_timestamp)
				.setBody('Second batched log record')
				.setEventName('BatchRecord2')
				.setStringAttribute('batch.position', 'second')
				.setNumberAttribute('batch.positionNum', _num)
				.emit(failureResult=>_loggerFailureResult);
			_num := 3;
			_thirdEmitSucceeded := _logger1
				.startLogRecord(severityNumber:=E_SeverityNumber.WARN)
				.setTimestamp(_timestamp)
				.setBody('Third batched log record')
				.setEventName('BatchRecord3')
				.setStringAttribute('batch.position', 'third')
				.setNumberAttribute('batch.positionNum', _num)
				.emit(failureResult=>_loggerFailureResult);
			_provider
				.stageProcessor(_processor)
				.tick();
			THIS^.AssertTrue(_firstEmitSucceeded, 'Expected the first emit to succeed');
			THIS^.AssertTrue(_secondEmitSucceeded, 'Expected the second emit to succeed');
			THIS^.AssertTrue(_thirdEmitSucceeded, 'Expected the third emit to succeed');
			THIS^.AssertTrue(_logger1.pLogRecord = 0, 'Expected emit to release the logger-owned record');
			IF _firstEmitSucceeded
				AND _secondEmitSucceeded
				AND _thirdEmitSucceeded THEN
				THIS^.AssertEquals_UDINT(3, _processor.records.count, 'Expected the processor to capture all three log records');
				_state := 10;
				RETURN;
			ELSE
				_state := 30;
				RETURN;
			END_IF
			
		10: // hand the captured records to the file exporter and tick it until the write is done
			IF _processor.records.count > 0 THEN
				_exportSucceeded := _processor.exportRecords(
					exporter:=_exporter,
					failureReason=>_exporterFailureReason
				);
				IF NOT _exportSucceeded OR_ELSE _processor.records.count > 0 THEN
					THIS^.AssertTrue(FALSE, 'Expected the exporter to take ownership of the processor buffer');
					_state := 30;
					RETURN;
				END_IF
			END_IF
			_exportCallSucceeded := _exporter.tick(failureReason=>_exporterFailureReason);
			_cycles := _cycles + 1;
			IF NOT _exportCallSucceeded THEN
				THIS^.AssertTrue(
					_exporterFailureReason <> E_LogRecordExporterFailureReason.NA,
					'Expected an exporter failure reason when tick returns FALSE'
				);
				THIS^.AssertTrue(FALSE, 'Expected the file export to succeed');
				_state := 30;
				RETURN;
			ELSIF _cycles > MAX_CYCLES THEN
				THIS^.AssertTrue(FALSE, 'Expected the file export to finish within MAX_CYCLES');
				_state := 30;
				RETURN;
			ELSIF _exporter.currentState = E_FileExporterState.done AND NOT _redelivered THEN
				// hand over the next batch in the same scan; the exporter must still start it
				_redelivered := TRUE;
				_logger2
					.startLogRecord(severityNumber:=E_SeverityNumber.INFO)
					.setTimestamp(_timestamp)
					.setBody('Batch exported the scan the previous one finished')
					.emit(failureResult=>_loggerFailureResult);
				_provider
					.stageProcessor(_processor)
					.tick();
				_exportSucceeded := _processor.exportRecords(
					exporter:=_exporter,
					failureReason=>_exporterFailureReason
				);
				THIS^.AssertTrue(_exportSucceeded, 'Expected the finished exporter to accept the next batch');
				RETURN;
			ELSIF _exporter.currentState = E_FileExporterState.done THEN
				THIS^.AssertFalse(_exporter.isBusy(), 'Expected the exporter to release its completed records');
				THIS^.AssertTrue(
					_exporterFailureReason = E_LogRecordExporterFailureReason.NA,
					'Expected no failure reason when file export succeeds'
				);
				_state := 20;
				RETURN;
			ELSE
				RETURN;
			END_IF
			
		20: // verify the exported batch made the file non-empty
			_fileFinder(
				sPathName:=_filepath,
				bExecute:=TRUE,
			);
			IF NOT _fileFinder.bBusy THEN
				_fileSize := ULARGE_TO_ULINT(_fileFinder.stFindFile.fileSize);
				THIS^.AssertTrue(_fileSize > 0, 'Expected a non-empty file');
				_state := 30;
			END_IF
			RETURN;
		
		30: // cleanup the file
			IF cleanup THEN
				_fileDeleter(
					sPathName:=_filepath,
					bExecute:=TRUE,
				);
				IF _fileDeleter.bBusy THEN
					RETURN;
				END_IF
			END_IF

			// clean up the record owned by the processor
			_processor.free();
			_logger1.free();
			THIS^.AssertTrue(_processor.records.count = 0, 'Expected the processor to be empty after cleanup');

			_state := 0;
			TcUnit.TEST_FINISHED();
	END_CASE
END_METHOD

END_FUNCTION_BLOCK

// ---- TEST/LOGGING/EXPORTING/FB_TestHttpExporter.TcPOU
(* Tests how the HTTP log exporter reports and recovers from destination failures. *)
FUNCTION_BLOCK FB_TestHttpExporter EXTENDS FB_TestSuite
VAR
	_exporterBadUrl: 	FB_LogRecordExporter_HTTP(url:='not-a-valid-url', bNoServerCertCheck:=TRUE);
	_exporterRefused: 	FB_LogRecordExporter_HTTP(url:='http://127.0.0.1:1/v1/logs', bNoServerCertCheck:=TRUE);
END_VAR

THIS^.testInvalidUrlFailsFast();
THIS^.testConnectionRefusedReportsFailure();

(*
	A refused connection surfaces as HTTP_REQUEST_FAILURE and leaves the exporter in the error state,
	and the next export still recovers it, so one unreachable collector cannot wedge logging for good.
*)
METHOD testConnectionRefusedReportsFailure : REFERENCE TO FB_Test

VAR CONSTANT
	MAX_CYCLES: UDINT := 60000;  // generous bound on scan cycles per request; a loopback refusal normally fails in a few
END_VAR

VAR_INST
	_cycles: 		UDINT;
	_state:			USINT;
END_VAR

VAR
	exportSucceeded: BOOL;
	callSucceeded: BOOL;
	failureReason: E_LogRecordExporterFailureReason;
END_VAR
TcUnit.TEST('testConnectionRefusedReportsFailure');
	CASE _state OF
		0: // export one batch to the unreachable endpoint
			_cycles := 0;
			exportSucceeded := THIS^._exportOneRecord(exporter:=_exporterRefused, timestamp:=1, failureReason=>failureReason);
			THIS^.AssertTrue(
				exportSucceeded
				AND_THEN failureReason = E_LogRecordExporterFailureReason.NA,
				'Expected the HTTP exporter to accept the batch for an unreachable endpoint'
			);
			_state := 10;
			RETURN;

		10: // wait for the request to fail; loopback refusal should be quick
			callSucceeded := _exporterRefused.tick(failureReason=>failureReason);
			_cycles := _cycles + 1;
			IF NOT callSucceeded THEN
				THIS^.AssertTrue(
					failureReason = E_LogRecordExporterFailureReason.HTTP_REQUEST_FAILURE,
					'Expected HTTP_REQUEST_FAILURE when the server refuses the connection'
				);
				THIS^.AssertTrue(
					_exporterRefused.currentState = E_HttpExporterState.error,
					'Expected the exporter to enter the error state after a refused connection'
				);
				_state := 15;
				RETURN;
			ELSIF _cycles > MAX_CYCLES THEN
				THIS^.AssertTrue(FALSE, 'Expected the refused connection to fail within MAX_CYCLES');
				_state := 20;
				RETURN;
			ELSE
				RETURN;
			END_IF

		15: // a failed export must not wedge the exporter; it accepts the next batch
			exportSucceeded := THIS^._exportOneRecord(exporter:=_exporterRefused, timestamp:=2, failureReason=>failureReason);
			THIS^.AssertTrue(
				exportSucceeded
				AND_THEN failureReason = E_LogRecordExporterFailureReason.NA
				AND_THEN _exporterRefused.currentState = E_HttpExporterState.idle,
				'Expected export to reset an errored exporter back to idle'
			);
			_cycles := 0;
			_state := 16;
			RETURN;

		16: // the accepted batch must start and fail again rather than wait in idle for good
			callSucceeded := _exporterRefused.tick(failureReason=>failureReason);
			_cycles := _cycles + 1;
			IF NOT callSucceeded THEN
				THIS^.AssertTrue(
					_exporterRefused.currentState = E_HttpExporterState.error,
					'Expected the second batch to reach the error state'
				);
				_state := 20;
			ELSIF _cycles > MAX_CYCLES THEN
				THIS^.AssertTrue(FALSE, CONCAT('Expected the second batch to fail within MAX_CYCLES; state ', TO_STRING(_exporterRefused.currentState)));
				_state := 20;
			END_IF
			RETURN;

		20: // cleanup
			_exporterRefused.free();
			THIS^.AssertFalse(_exporterRefused.isBusy(), 'Expected the HTTP exporter to release its records on cleanup');
			_state := 0;
			TcUnit.TEST_FINISHED();
	END_CASE
END_METHOD

(*
	An endpoint URL without an http(s) scheme fails on the first tick with HTTP_URL_PARSE_FAILURE and
	releases the batch without sending, so a misconfigured exporter never holds records or blocks a request slot.
*)
METHOD testInvalidUrlFailsFast : REFERENCE TO FB_Test
VAR
	exportSucceeded: BOOL;
	callSucceeded: BOOL;
	failureReason: E_LogRecordExporterFailureReason;
END_VAR
TcUnit.TEST('testInvalidUrlFailsFast');
	exportSucceeded := THIS^._exportOneRecord(exporter:=_exporterBadUrl, timestamp:=1, failureReason=>failureReason);
	THIS^.AssertTrue(
		exportSucceeded
		AND_THEN failureReason = E_LogRecordExporterFailureReason.NA,
		'Expected the exporter to accept the batch before validating the URL'
	);

	callSucceeded := _exporterBadUrl.tick(failureReason=>failureReason);
	THIS^.AssertFalse(callSucceeded, 'Expected tick to report failure for an unparseable endpoint URL');
	THIS^.AssertTrue(
		failureReason = E_LogRecordExporterFailureReason.HTTP_URL_PARSE_FAILURE,
		'Expected HTTP_URL_PARSE_FAILURE for an endpoint URL without an http(s) scheme'
	);
	THIS^.AssertTrue(
		_exporterBadUrl.currentState = E_HttpExporterState.error,
		'Expected the exporter to enter the error state without sending anything'
	);
	THIS^.AssertFalse(_exporterBadUrl.isBusy(), 'Expected the failed batch to be released');

	// A failed exporter recovers when the next export is accepted.
	exportSucceeded := THIS^._exportOneRecord(exporter:=_exporterBadUrl, timestamp:=2, failureReason=>failureReason);
	THIS^.AssertTrue(
		exportSucceeded
		AND_THEN _exporterBadUrl.currentState = E_HttpExporterState.idle,
		'Expected export to reset an errored exporter back to idle'
	);

	_exporterBadUrl.free();
TcUnit.TEST_FINISHED();
END_METHOD

(*
	Emits one record through a logger and hands it to the exporter as a one-record batch,
	asserting that the record reached the batch and that the exporter took it out.
	Returns what export returned.
*)
METHOD _exportOneRecord : BOOL
VAR_INPUT
	exporter: REFERENCE TO FB_LogRecordExporter_Base;
	timestamp: ULINT;
END_VAR
VAR_OUTPUT
	failureReason: E_LogRecordExporterFailureReason;
END_VAR
VAR
	resource: FB_Resource(schemaUrl:='');
	provider: FB_LoggerProvider(resource:=resource);
	scope: FB_InstrumentationScope(name:='http.exporter.test', version:='1.0.0', schemaUrl:='');
	logger: FB_Logger(scope:=scope, provider:=provider);
	processor: FB_LogRecordProcessor_ForRecordsInspection(
		maxQueueSize:=0,
		scheduledDelayMillis:=1000,
		maxExportBatchSize:=512,
		exporter:=0
	);
	emitSucceeded: BOOL;
	emitFailureReason: E_LoggerFailureReason;
END_VAR
_exportOneRecord := FALSE;
emitSucceeded := logger
	.startLogRecord(severityNumber:=E_SeverityNumber.INFO)
	.setTimestamp(timestamp)
	.emit(failureResult=>emitFailureReason);
provider
	.stageProcessor(processor)
	.tick();
THIS^.AssertTrue(emitSucceeded AND_THEN processor.records.count = 1, 'Expected the logger to hand one record to the batch');

_exportOneRecord := processor.exportRecords(exporter:=exporter, failureReason=>failureReason);
THIS^.AssertEquals_UDINT(0, processor.records.count, 'Expected the exporter to take the record out of the batch');
processor.free();
END_METHOD

END_FUNCTION_BLOCK

// ---- TEST/TRACING/ID_GENERATOR/FB_TestIdGenerator.TcPOU
(* Tests trace and span identifier generation.

   A generator fills its ring from the operating system guid service over ADS, so a fresh one
   has nothing to hand out until tick has been pumped for a few cycles. Every test that needs
   identifiers waits for that first refill before asserting anything about the bytes it gets
   back.

   Each test declares its generator in its own VAR_INST, next to the state machine that pumps
   it, so the ring a test reasons about is written down where the test reads it rather than in
   a list on the suite. Ring sizes are therefore chosen per test: most take a ring far larger
   than they draw from, so the seam never comes into it, while the wrap and capacity tests
   deliberately take the smallest ring the configuration allows, because a ring that small is
   the only one a test can drain often enough to lap. *)
FUNCTION_BLOCK FB_TestIdGenerator EXTENDS FB_TestSuite

THIS^.testRejectsInvalidConfiguration();
THIS^.testFailsBeforeTheFirstRefill();
THIS^.testGeneratesUniqueTraceIds();
THIS^.testGeneratesUniqueSpanIds();
THIS^.testDrawsAcrossTheWrap();
THIS^.testHonorsConfiguredCapacity();
THIS^.testGeneratesThroughTheBaseReference();
THIS^.testSeparateGeneratorsDoNotCollide();

(* TRUE when every byte in the buffer is zero, which is the identifier OTLP reads as absent. *)
METHOD _isZero : BOOL
VAR_INPUT
	pBytes: POINTER TO BYTE;
	nBytes: UDINT;
END_VAR
VAR
	_idx: UDINT;
END_VAR
_isZero := TRUE;

IF (pBytes = 0) OR_ELSE (nBytes = 0) THEN
	RETURN;
END_IF

FOR _idx := 0 TO nBytes - 1 DO
	IF pBytes[_idx] <> 0 THEN
		_isZero := FALSE;
		RETURN;
	END_IF
END_FOR
END_METHOD

(* Exercises the seam. A thirty two byte ring cannot hold eight identifiers at once, so the
   draws are spread over cycles and the read point laps the ring several times.

   Taking sixteen bytes and then eight moves the read point by twenty four, which lands it on
   every eight byte alignment in turn: some trace draws stop short of the end of the ring, one
   ends exactly on it, and one starts near the end and has to be stitched from both sides. A
   stitch that copied the wrong end, or re-read bytes already handed out, shows up here as a
   repeat among the samples. *)
METHOD testDrawsAcrossTheWrap : REFERENCE TO FB_Test

VAR CONSTANT
	MAX_CYCLES: UDINT := 60000;
	SAMPLES: UDINT := 8;
END_VAR

VAR_INST
	_generator: FB_IdGenerator(nTraceIds := 1, nSpanIds := 1);  // 24 bytes, which FB_Init rounds up to 32
	_cycles: UDINT;
	_state: USINT;
	_traceIdx: UDINT;
	_spanIdx: UDINT;
	_traceSamples: ARRAY [0..7, 0..15] OF BYTE;  // held across cycles, unlike the other suites
	_spanSamples: ARRAY [0..7, 0..7] OF BYTE;
END_VAR

VAR
	traceId: FB_TraceId;
	spanId: FB_SpanId;
	failureReason: E_IdGenFailureReason;
	tickSucceeded: BOOL;
	_i: UDINT;
	_j: UDINT;
END_VAR
TcUnit.TEST('testDrawsAcrossTheWrap');
	CASE _state OF
		0: // take whatever the ring can serve this cycle, however many laps that takes
			tickSucceeded := _generator.tick(failureReason=>failureReason);
			_cycles := _cycles + 1;
			IF NOT tickSucceeded THEN
				THIS^.AssertTrue(FALSE, 'Expected the guid service to refill the ring without error');
				_state := 255;
				TcUnit.TEST_FINISHED();
				RETURN;
			END_IF

			IF (_traceIdx < SAMPLES) AND_THEN _generator.generateTraceId(traceId:=traceId, failureReason=>failureReason) THEN
				MEMCPY(ADR(_traceSamples[_traceIdx, 0]), ADR(traceId.bytes), SIZEOF(traceId.bytes));
				_traceIdx := _traceIdx + 1;
			END_IF

			IF (_spanIdx < SAMPLES) AND_THEN _generator.generateSpanId(spanId:=spanId, failureReason=>failureReason) THEN
				MEMCPY(ADR(_spanSamples[_spanIdx, 0]), ADR(spanId.bytes), SIZEOF(spanId.bytes));
				_spanIdx := _spanIdx + 1;
			END_IF

			IF (_traceIdx >= SAMPLES) AND (_spanIdx >= SAMPLES) THEN
				_state := 10;
			ELSIF _cycles > MAX_CYCLES THEN
				THIS^.AssertTrue(FALSE, 'Expected a ring small enough to wrap to hand out its identifiers within MAX_CYCLES');
				_state := 255;
				TcUnit.TEST_FINISHED();
			END_IF
			RETURN;

		10:
			FOR _i := 0 TO 7 DO
				THIS^.AssertFalse(
					THIS^._isZero(pBytes:=ADR(_traceSamples[_i, 0]), nBytes:=TO_UDINT(SIZEOF(traceId.bytes))),
					'Expected no trace id drawn from a wrapping ring to be all zeroes'
				);
				THIS^.AssertFalse(
					THIS^._isZero(pBytes:=ADR(_spanSamples[_i, 0]), nBytes:=TO_UDINT(SIZEOF(spanId.bytes))),
					'Expected no span id drawn from a wrapping ring to be all zeroes'
				);

				FOR _j := 0 TO 7 DO
					IF _i <> _j THEN
						THIS^.AssertTrue(
							MEMCMP(ADR(_traceSamples[_i, 0]), ADR(_traceSamples[_j, 0]), SIZEOF(traceId.bytes)) <> 0,
							'Expected every trace id to differ, including the one stitched across the wrap'
						);
						THIS^.AssertTrue(
							MEMCMP(ADR(_spanSamples[_i, 0]), ADR(_spanSamples[_j, 0]), SIZEOF(spanId.bytes)) <> 0,
							'Expected every span id to differ, including the ones taken either side of the wrap'
						);
					END_IF
				END_FOR
			END_FOR

			_state := 255;
			TcUnit.TEST_FINISHED();
			RETURN;
	END_CASE
END_METHOD

(* A generator that has never been ticked holds no bytes. It has to say so, because the only
   thing it could hand out instead is the all zero identifier OTLP reads as absent. *)
METHOD testFailsBeforeTheFirstRefill : REFERENCE TO FB_Test

VAR_INST
	_generator: FB_IdGenerator(nTraceIds := 16, nSpanIds := 16);  // deliberately never ticked, so it stays empty
	_state: USINT;
END_VAR

VAR
	traceId: FB_TraceId;
	spanId: FB_SpanId;
	failureReason: E_IdGenFailureReason;
	success: BOOL;
END_VAR
TcUnit.TEST('testFailsBeforeTheFirstRefill');
	CASE _state OF
		0:
			THIS^.AssertTrue(_generator.configValid, 'Expected a generator with a ring to report a valid configuration');

			success := _generator.generateTraceId(traceId:=traceId, failureReason=>failureReason);
			THIS^.AssertFalse(success, 'Expected trace id generation to fail before the first refill');
			THIS^.AssertEquals_UDINT(
				TO_UDINT(E_IdGenFailureReason.NO_IDENTIFIERS_AVAILABLE),
				TO_UDINT(failureReason),
				'Expected an empty ring to report NO_IDENTIFIERS_AVAILABLE'
			);
			THIS^.AssertTrue(
				THIS^._isZero(pBytes:=ADR(traceId.bytes), nBytes:=TO_UDINT(SIZEOF(traceId.bytes))),
				'Expected a failed draw to leave the trace id untouched'
			);

			success := _generator.generateSpanId(spanId:=spanId, failureReason=>failureReason);
			THIS^.AssertFalse(success, 'Expected span id generation to fail before the first refill');
			THIS^.AssertEquals_UDINT(
				TO_UDINT(E_IdGenFailureReason.NO_IDENTIFIERS_AVAILABLE),
				TO_UDINT(failureReason),
				'Expected an empty ring to report NO_IDENTIFIERS_AVAILABLE'
			);
			THIS^.AssertTrue(
				THIS^._isZero(pBytes:=ADR(spanId.bytes), nBytes:=TO_UDINT(SIZEOF(spanId.bytes))),
				'Expected a failed draw to leave the span id untouched'
			);

			_state := 255;
			TcUnit.TEST_FINISHED();
	END_CASE
END_METHOD

(* Callers hold the generator as REFERENCE TO FB_IdGenerator_Base, so the abstract methods have
   to dispatch to the concrete ring. *)
METHOD testGeneratesThroughTheBaseReference : REFERENCE TO FB_Test

VAR CONSTANT
	MAX_CYCLES: UDINT := 60000;
END_VAR

VAR_INST
	_generator: FB_IdGenerator(nTraceIds := 16, nSpanIds := 16);
	_cycles: UDINT;
	_state: USINT;
END_VAR

VAR
	base: REFERENCE TO FB_IdGenerator_Base;
	traceId: FB_TraceId;
	spanId: FB_SpanId;
	failureReason: E_IdGenFailureReason;
	tickSucceeded: BOOL;
	success: BOOL;
END_VAR
TcUnit.TEST('testGeneratesThroughTheBaseReference');
	base REF= _generator;
	CASE _state OF
		0:
			THIS^.AssertTrue(__ISVALIDREF(base), 'Expected the base reference to be valid');
			_state := 10;
			RETURN;

		10: // pump through the base reference until the first refill lands
			tickSucceeded := base.tick(failureReason=>failureReason);
			_cycles := _cycles + 1;
			IF NOT tickSucceeded THEN
				THIS^.AssertTrue(FALSE, 'Expected tick to dispatch to the concrete generator without error');
				_state := 255;
				TcUnit.TEST_FINISHED();
				RETURN;
			END_IF

			success := base.generateTraceId(traceId:=traceId, failureReason=>failureReason);
			IF NOT success THEN
				IF _cycles > MAX_CYCLES THEN
					THIS^.AssertTrue(FALSE, 'Expected identifiers through the base reference within MAX_CYCLES');
					_state := 255;
					TcUnit.TEST_FINISHED();
				END_IF
				RETURN;
			END_IF

			THIS^.AssertFalse(
				THIS^._isZero(pBytes:=ADR(traceId.bytes), nBytes:=TO_UDINT(SIZEOF(traceId.bytes))),
				'Expected a non zero trace id through the base reference'
			);

			success := base.generateSpanId(spanId:=spanId, failureReason=>failureReason);
			THIS^.AssertTrue(success, 'Expected generateSpanId to dispatch to the concrete generator');
			THIS^.AssertFalse(
				THIS^._isZero(pBytes:=ADR(spanId.bytes), nBytes:=TO_UDINT(SIZEOF(spanId.bytes))),
				'Expected a non zero span id through the base reference'
			);

			_state := 255;
			TcUnit.TEST_FINISHED();
			RETURN;
	END_CASE
END_METHOD

(* The same requirement as for trace ids. A span id handed out twice makes two spans in the
   same trace indistinguishable. *)
METHOD testGeneratesUniqueSpanIds : REFERENCE TO FB_Test

VAR CONSTANT
	MAX_CYCLES: UDINT := 60000;
END_VAR

VAR_INST
	_generator: FB_IdGenerator(nTraceIds := 16, nSpanIds := 16);  // 384 bytes, so eight samples come out of one fill
	_cycles: UDINT;
	_state: USINT;
END_VAR

VAR
	spanId: FB_SpanId;
	samples: ARRAY [0..7, 0..7] OF BYTE;
	failureReason: E_IdGenFailureReason;
	tickSucceeded: BOOL;
	success: BOOL;
	_i: UDINT;
	_j: UDINT;
END_VAR
TcUnit.TEST('testGeneratesUniqueSpanIds');
	CASE _state OF
		0: // wait for the first refill before drawing the samples
			tickSucceeded := _generator.tick(failureReason=>failureReason);
			_cycles := _cycles + 1;
			IF NOT tickSucceeded THEN
				THIS^.AssertTrue(FALSE, 'Expected the guid service to refill the ring without error');
				_state := 255;
				TcUnit.TEST_FINISHED();
				RETURN;
			END_IF

			IF _generator.generateSpanId(spanId:=spanId, failureReason=>failureReason) THEN
				_state := 10;
			ELSIF _cycles > MAX_CYCLES THEN
				THIS^.AssertTrue(FALSE, 'Expected the first ring of span ids within MAX_CYCLES');
				_state := 255;
				TcUnit.TEST_FINISHED();
			END_IF
			RETURN;

		10: // a full ring holds forty eight span ids, so all eight samples come out of one fill
			FOR _i := 0 TO 7 DO
				success := _generator.generateSpanId(spanId:=spanId, failureReason=>failureReason);
				THIS^.AssertTrue(success, 'Expected every span id draw from a filled ring to succeed');
				THIS^.AssertEquals_UDINT(
					TO_UDINT(E_IdGenFailureReason.NA),
					TO_UDINT(failureReason),
					'Expected no failure reason alongside a successful draw'
				);
				THIS^.AssertFalse(
					THIS^._isZero(pBytes:=ADR(spanId.bytes), nBytes:=TO_UDINT(SIZEOF(spanId.bytes))),
					'Expected no span id to be all zeroes'
				);
				MEMCPY(ADR(samples[_i, 0]), ADR(spanId.bytes), SIZEOF(spanId.bytes));
			END_FOR

			FOR _i := 0 TO 7 DO
				FOR _j := 0 TO 7 DO
					IF _i <> _j THEN
						THIS^.AssertTrue(
							MEMCMP(ADR(samples[_i, 0]), ADR(samples[_j, 0]), SIZEOF(spanId.bytes)) <> 0,
							'Expected every span id to differ from every other'
						);
					END_IF
				END_FOR
			END_FOR

			_state := 255;
			TcUnit.TEST_FINISHED();
			RETURN;
	END_CASE
END_METHOD

(* Every draw has to be its own bytes. A trace id handed out twice merges two unrelated traces
   at the collector, which is worse than no trace at all. *)
METHOD testGeneratesUniqueTraceIds : REFERENCE TO FB_Test

VAR CONSTANT
	MAX_CYCLES: UDINT := 60000;
END_VAR

VAR_INST
	_generator: FB_IdGenerator(nTraceIds := 16, nSpanIds := 16);  // 384 bytes, so eight samples come out of one fill
	_cycles: UDINT;
	_state: USINT;
END_VAR

VAR
	traceId: FB_TraceId;
	samples: ARRAY [0..7, 0..15] OF BYTE;
	failureReason: E_IdGenFailureReason;
	tickSucceeded: BOOL;
	success: BOOL;
	_i: UDINT;
	_j: UDINT;
END_VAR
TcUnit.TEST('testGeneratesUniqueTraceIds');
	CASE _state OF
		0: // wait for the first refill before drawing the samples
			tickSucceeded := _generator.tick(failureReason=>failureReason);
			_cycles := _cycles + 1;
			IF NOT tickSucceeded THEN
				THIS^.AssertTrue(FALSE, 'Expected the guid service to refill the ring without error');
				_state := 255;
				TcUnit.TEST_FINISHED();
				RETURN;
			END_IF

			IF _generator.generateTraceId(traceId:=traceId, failureReason=>failureReason) THEN
				_state := 10;
			ELSIF _cycles > MAX_CYCLES THEN
				THIS^.AssertTrue(FALSE, 'Expected the first ring of trace ids within MAX_CYCLES');
				_state := 255;
				TcUnit.TEST_FINISHED();
			END_IF
			RETURN;

		10: // a full ring holds twenty four trace ids, so all eight samples come out of one fill
			FOR _i := 0 TO 7 DO
				success := _generator.generateTraceId(traceId:=traceId, failureReason=>failureReason);
				THIS^.AssertTrue(success, 'Expected every trace id draw from a filled ring to succeed');
				THIS^.AssertEquals_UDINT(
					TO_UDINT(E_IdGenFailureReason.NA),
					TO_UDINT(failureReason),
					'Expected no failure reason alongside a successful draw'
				);
				THIS^.AssertFalse(
					THIS^._isZero(pBytes:=ADR(traceId.bytes), nBytes:=TO_UDINT(SIZEOF(traceId.bytes))),
					'Expected no trace id to be all zeroes'
				);
				MEMCPY(ADR(samples[_i, 0]), ADR(traceId.bytes), SIZEOF(traceId.bytes));
			END_FOR

			FOR _i := 0 TO 7 DO
				FOR _j := 0 TO 7 DO
					IF _i <> _j THEN
						THIS^.AssertTrue(
							MEMCMP(ADR(samples[_i, 0]), ADR(samples[_j, 0]), SIZEOF(traceId.bytes)) <> 0,
							'Expected every trace id to differ from every other'
						);
					END_IF
				END_FOR
			END_FOR

			_state := 255;
			TcUnit.TEST_FINISHED();
			RETURN;
	END_CASE
END_METHOD

(* One trace id and one span id is twenty four bytes, which FB_Init rounds up to thirty two
   because the guid service will not write anything narrower than a whole guid. A full ring is
   therefore exactly two trace ids wide, and no amount of refilling grows it past that. *)
METHOD testHonorsConfiguredCapacity : REFERENCE TO FB_Test

VAR CONSTANT
	MAX_CYCLES: UDINT := 60000;
	MAX_DRAWS: UDINT := 16;  // comfortably more than a thirty two byte ring could ever serve
	EXPECTED_TRACE_IDS: UDINT := 2;
END_VAR

VAR_INST
	_generator: FB_IdGenerator(nTraceIds := 1, nSpanIds := 1);  // the shortest ring the configuration allows
	_cycles: UDINT;
	_state: USINT;
	_best: UDINT;  // the most trace ids any single drain has yielded
END_VAR

VAR
	traceId: FB_TraceId;
	failureReason: E_IdGenFailureReason;
	tickSucceeded: BOOL;
	drawn: UDINT;
	_i: UDINT;
END_VAR
TcUnit.TEST('testHonorsConfiguredCapacity');
	CASE _state OF
		0: // drain the ring dry every cycle, so the best any one drain manages is one full ring
			tickSucceeded := _generator.tick(failureReason=>failureReason);
			_cycles := _cycles + 1;
			IF NOT tickSucceeded THEN
				THIS^.AssertTrue(FALSE, 'Expected the guid service to refill the ring without error');
				_state := 255;
				TcUnit.TEST_FINISHED();
				RETURN;
			END_IF

			drawn := 0;
			FOR _i := 1 TO MAX_DRAWS DO
				IF NOT _generator.generateTraceId(traceId:=traceId, failureReason=>failureReason) THEN
					EXIT;
				END_IF
				drawn := drawn + 1;
			END_FOR

			THIS^.AssertTrue(
				drawn <= EXPECTED_TRACE_IDS,
				'Expected a refill never to serve more than the configured ring holds'
			);
			THIS^.AssertEquals_UDINT(
				TO_UDINT(E_IdGenFailureReason.NO_IDENTIFIERS_AVAILABLE),
				TO_UDINT(failureReason),
				'Expected the draw that emptied the ring to report NO_IDENTIFIERS_AVAILABLE'
			);

			IF drawn > _best THEN
				_best := drawn;
			END_IF

			IF _best >= EXPECTED_TRACE_IDS THEN
				_state := 10;
			ELSIF _cycles > MAX_CYCLES THEN
				THIS^.AssertTrue(FALSE, 'Expected the ring to fill to its configured length within MAX_CYCLES');
				_state := 255;
				TcUnit.TEST_FINISHED();
			END_IF
			RETURN;

		10:
			THIS^.AssertEquals_UDINT(
				EXPECTED_TRACE_IDS,
				_best,
				'Expected a twenty four byte request to become a thirty two byte ring'
			);
			_state := 255;
			TcUnit.TEST_FINISHED();
			RETURN;
	END_CASE
END_METHOD

(* A generator asked for no identifiers never allocates a ring, so every entry point has to say
   so rather than read through a null pointer. *)
METHOD testRejectsInvalidConfiguration : REFERENCE TO FB_Test

VAR_INST
	_generator: FB_IdGenerator(nTraceIds := 0, nSpanIds := 0);  // asks for nothing, so no ring is allocated
	_state: USINT;
END_VAR

VAR
	traceId: FB_TraceId;
	spanId: FB_SpanId;
	failureReason: E_IdGenFailureReason;
	success: BOOL;
END_VAR
TcUnit.TEST('testRejectsInvalidConfiguration');
	CASE _state OF
		0:
			THIS^.AssertFalse(_generator.configValid, 'Expected a generator with no ring to report an invalid configuration');

			success := _generator.tick(failureReason=>failureReason);
			THIS^.AssertFalse(success, 'Expected tick to fail when no ring was allocated');
			THIS^.AssertEquals_UDINT(
				TO_UDINT(E_IdGenFailureReason.INVALID_CONFIGUATION),
				TO_UDINT(failureReason),
				'Expected tick to report INVALID_CONFIGUATION'
			);

			success := _generator.generateTraceId(traceId:=traceId, failureReason=>failureReason);
			THIS^.AssertFalse(success, 'Expected trace id generation to fail when no ring was allocated');
			THIS^.AssertEquals_UDINT(
				TO_UDINT(E_IdGenFailureReason.INVALID_CONFIGUATION),
				TO_UDINT(failureReason),
				'Expected a missing ring to be reported as a configuration mistake, not an empty ring'
			);

			success := _generator.generateSpanId(spanId:=spanId, failureReason=>failureReason);
			THIS^.AssertFalse(success, 'Expected span id generation to fail when no ring was allocated');
			THIS^.AssertEquals_UDINT(
				TO_UDINT(E_IdGenFailureReason.INVALID_CONFIGUATION),
				TO_UDINT(failureReason),
				'Expected a missing ring to be reported as a configuration mistake, not an empty ring'
			);

			_state := 255;
			TcUnit.TEST_FINISHED();
	END_CASE
END_METHOD

(* Two generators built in the same cycle must not emit the same identifiers, or two providers
   on one PLC would report traces the collector cannot tell apart. *)
METHOD testSeparateGeneratorsDoNotCollide : REFERENCE TO FB_Test

VAR CONSTANT
	MAX_CYCLES: UDINT := 60000;
END_VAR

VAR_INST
	_generatorA: FB_IdGenerator(nTraceIds := 16, nSpanIds := 16);
	_generatorB: FB_IdGenerator(nTraceIds := 16, nSpanIds := 16);
	_cycles: UDINT;
	_state: USINT;
END_VAR

VAR
	traceIdA: FB_TraceId;
	traceIdB: FB_TraceId;
	spanIdA: FB_SpanId;
	spanIdB: FB_SpanId;
	failureReason: E_IdGenFailureReason;
	tickSucceededA: BOOL;
	tickSucceededB: BOOL;
	drewA: BOOL;
	drewB: BOOL;
	success: BOOL;
END_VAR
TcUnit.TEST('testSeparateGeneratorsDoNotCollide');
	CASE _state OF
		0: // pump both rings until they can each serve in the same cycle
			tickSucceededA := _generatorA.tick(failureReason=>failureReason);
			tickSucceededB := _generatorB.tick(failureReason=>failureReason);
			_cycles := _cycles + 1;
			IF NOT (tickSucceededA AND tickSucceededB) THEN
				THIS^.AssertTrue(FALSE, 'Expected both generators to refill without error');
				_state := 255;
				TcUnit.TEST_FINISHED();
				RETURN;
			END_IF

			// both are drawn unconditionally, so neither ring is drained ahead of the other
			drewA := _generatorA.generateTraceId(traceId:=traceIdA, failureReason=>failureReason);
			drewB := _generatorB.generateTraceId(traceId:=traceIdB, failureReason=>failureReason);
			IF NOT (drewA AND drewB) THEN
				IF _cycles > MAX_CYCLES THEN
					THIS^.AssertTrue(FALSE, 'Expected both generators to fill within MAX_CYCLES');
					_state := 255;
					TcUnit.TEST_FINISHED();
				END_IF
				RETURN;
			END_IF

			THIS^.AssertTrue(
				MEMCMP(ADR(traceIdA.bytes), ADR(traceIdB.bytes), SIZEOF(traceIdA.bytes)) <> 0,
				'Expected two generators to produce different trace ids'
			);

			success := _generatorA.generateSpanId(spanId:=spanIdA, failureReason=>failureReason);
			THIS^.AssertTrue(success, 'Expected the first generator to serve a span id from a filled ring');
			success := _generatorB.generateSpanId(spanId:=spanIdB, failureReason=>failureReason);
			THIS^.AssertTrue(success, 'Expected the second generator to serve a span id from a filled ring');
			THIS^.AssertTrue(
				MEMCMP(ADR(spanIdA.bytes), ADR(spanIdB.bytes), SIZEOF(spanIdA.bytes)) <> 0,
				'Expected two generators to produce different span ids'
			);

			_state := 255;
			TcUnit.TEST_FINISHED();
			RETURN;
	END_CASE
END_METHOD

END_FUNCTION_BLOCK

// ---- TEST/TRACING/SPAN/FB_TestSpanContext.TcPOU
(* Tests the span context value object and ContextFactory.buildContext and fromSpan: that a context holds
   copies of what it is built from, does not validate its identity, decodes remoteness from both
   flag bits, and releases its trace state.

   Every test deletes the contexts it builds before returning. *)
FUNCTION_BLOCK FB_TestSpanContext EXTENDS FB_TestSuite

THIS^.testBuildsCopiesOfItsInputs();
THIS^.testBuildsWithoutTraceState();
THIS^.testBuildsFromZeroIdentifiers();
THIS^.testRejectsAssignedDestination();
THIS^.testRejectsNullIdentifiers();
THIS^.testFromSpanRejectsNullSpan();
THIS^.testIsRemoteNeedsBothBits();
THIS^.testFreeClearsTheContext();
THIS^.testDeleteClearsTheCallersPointer();
THIS^.testDeleteRefusesAnotherPointer();

(* Writes distinct non-zero bytes into both identifiers, offset by seed so two calls with
   different seeds produce identifiers that can be told apart. *)
METHOD _fillIds
VAR_IN_OUT
	traceId: FB_TraceId;
	spanId: FB_SpanId;
END_VAR
VAR_INPUT
	seed: BYTE;
END_VAR
VAR
	_idx: UDINT;
	_bytes: ARRAY [0..15] OF BYTE;
END_VAR
// the identifier bytes are outputs, so they are written through their address
FOR _idx := 0 TO SIZEOF(_bytes) - 1 DO
	_bytes[_idx] := seed + TO_BYTE(_idx) + 1;
END_FOR
MEMCPY(ADR(traceId.bytes), ADR(_bytes), SIZEOF(traceId.bytes));

FOR _idx := 0 TO SIZEOF(_bytes) - 1 DO
	_bytes[_idx] := seed + TO_BYTE(_idx) + 16#40;
END_FOR
MEMCPY(ADR(spanId.bytes), ADR(_bytes), SIZEOF(spanId.bytes));
END_METHOD

(* Deletes a context built by a test and clears the pointer. *)
METHOD _release
VAR_IN_OUT
	pContext: POINTER TO FB_SpanContext;
END_VAR
IF pContext <> 0 THEN
	pContext^.delete(pSelf:=pContext);
END_IF
END_METHOD

(* A context outlives the span it came from, so it must hold copies. Changing the source
   identifiers or trace state after building must not change the context. *)
METHOD testBuildsCopiesOfItsInputs : REFERENCE TO FB_Test
VAR
	pContext: POINTER TO FB_SpanContext;
	traceId: FB_TraceId;
	spanId: FB_SpanId;
	expectedTraceId: FB_TraceId;
	expectedSpanId: FB_SpanId;
	traceState: T_MaxString := 'vendor=abc';
	pTraceState: POINTER TO FB_TraceState;
	success: BOOL;
	failureReason: E_ContextFactoryFailureReason;
END_VAR
TcUnit.TEST('testBuildsCopiesOfItsInputs');
	TraceStateFactory.parse(pDest:=pTraceState, pHeader:=ADR(traceState));
	THIS^._fillIds(traceId:=traceId, spanId:=spanId, seed:=0);
	THIS^._fillIds(traceId:=expectedTraceId, spanId:=expectedSpanId, seed:=0);

	success := ContextFactory.buildContext(
		pDest:=pContext,
		pTraceId:=ADR(traceId),
		pSpanId:=ADR(spanId),
		pTraceState:=pTraceState,
		traceFlags:=1,  // sampled
		failureReason=>failureReason
	);
	// the trace state is borrowed, so the caller releases its own copy at once
	IF pTraceState <> 0 THEN pTraceState^.delete(pSelf:=pTraceState); END_IF
	THIS^.AssertTrue(success, 'Expected buildContext to succeed');
	THIS^.AssertEquals_UDINT(
		TO_UDINT(E_ContextFactoryFailureReason.NA),
		TO_UDINT(failureReason),
		'Expected no failure reason on success'
	);
	THIS^.AssertTrue(pContext <> 0, 'Expected buildContext to assign the destination');
	IF pContext = 0 THEN
		TcUnit.TEST_FINISHED();
		RETURN;
	END_IF
	THIS^.AssertTrue(pContext^.isValid(), 'Expected a context built from non-zero identifiers to be valid');
	THIS^.AssertEquals_UDINT(1, pContext^.traceFlags, 'Expected the trace flags to be stored as given');

	// change every source after the fact
	THIS^._fillIds(traceId:=traceId, spanId:=spanId, seed:=16#80);

	THIS^.AssertTrue(
		MEMCMP(ADR(pContext^.traceId.bytes), ADR(expectedTraceId.bytes), SIZEOF(expectedTraceId.bytes)) = 0,
		'Expected the trace id to be a copy that does not follow its source'
	);
	THIS^.AssertTrue(
		MEMCMP(ADR(pContext^.spanId.bytes), ADR(expectedSpanId.bytes), SIZEOF(expectedSpanId.bytes)) = 0,
		'Expected the span id to be a copy that does not follow its source'
	);
	THIS^.AssertTrue(pContext^.traceState <> 0, 'Expected the trace state to be stored');
	IF pContext^.traceState <> 0 THEN
		THIS^.AssertEquals_STRING('vendor=abc', pContext^.traceState^.pString^, 'Expected the trace state to outlive its source');
	END_IF

	THIS^._release(pContext:=pContext);
TcUnit.TEST_FINISHED();
END_METHOD

(* Validation belongs to the producers of a context, not to the factory. All-zero identifiers
   build a context that exists but reports itself as not valid. *)
METHOD testBuildsFromZeroIdentifiers : REFERENCE TO FB_Test
VAR
	pContext: POINTER TO FB_SpanContext;
	zeroTraceId: FB_TraceId;
	zeroSpanId: FB_SpanId;
	success: BOOL;
	failureReason: E_ContextFactoryFailureReason;
END_VAR
TcUnit.TEST('testBuildsFromZeroIdentifiers');
	success := ContextFactory.buildContext(
		pDest:=pContext,
		pTraceId:=ADR(zeroTraceId),
		pSpanId:=ADR(zeroSpanId),
		pTraceState:=0,
		traceFlags:=0,
		failureReason=>failureReason
	);
	THIS^.AssertTrue(success, 'Expected buildContext not to validate the identifiers');
	THIS^.AssertEquals_UDINT(
		TO_UDINT(E_ContextFactoryFailureReason.NA),
		TO_UDINT(failureReason),
		'Expected no failure reason for all-zero identifiers'
	);
	THIS^.AssertTrue(pContext <> 0, 'Expected buildContext to assign the destination');
	IF pContext <> 0 THEN
		THIS^.AssertFalse(pContext^.isValid(), 'Expected a context with all-zero identifiers to be invalid');
		THIS^.AssertFalse(pContext^.isRemote(), 'Expected a context without remote bits not to report remote');
	END_IF

	THIS^._release(pContext:=pContext);
TcUnit.TEST_FINISHED();
END_METHOD

(* Trace state is optional; a null pointer means the context carries none. *)
METHOD testBuildsWithoutTraceState : REFERENCE TO FB_Test
VAR
	pContext: POINTER TO FB_SpanContext;
	traceId: FB_TraceId;
	spanId: FB_SpanId;
	success: BOOL;
	failureReason: E_ContextFactoryFailureReason;
END_VAR
TcUnit.TEST('testBuildsWithoutTraceState');
	THIS^._fillIds(traceId:=traceId, spanId:=spanId, seed:=0);

	success := ContextFactory.buildContext(
		pDest:=pContext,
		pTraceId:=ADR(traceId),
		pSpanId:=ADR(spanId),
		pTraceState:=0,
		traceFlags:=0,
		failureReason=>failureReason
	);
	THIS^.AssertTrue(success, 'Expected buildContext to succeed without a trace state');
	THIS^.AssertTrue(pContext <> 0, 'Expected buildContext to assign the destination');
	IF pContext <> 0 THEN
		THIS^.AssertTrue(pContext^.isValid(), 'Expected the context to be valid');
		THIS^.AssertTrue(pContext^.traceState = 0, 'Expected no trace state to be stored');
	END_IF

	THIS^._release(pContext:=pContext);
TcUnit.TEST_FINISHED();
END_METHOD

(* delete takes the caller's pointer by reference and clears it, so a released context can
   never be reached through the pointer that owned it. *)
METHOD testDeleteClearsTheCallersPointer : REFERENCE TO FB_Test
VAR
	pContext: POINTER TO FB_SpanContext;
	traceId: FB_TraceId;
	spanId: FB_SpanId;
	traceState: T_MaxString := 'vendor=abc';
	pTraceState: POINTER TO FB_TraceState;
	deleted: BOOL;
END_VAR
TcUnit.TEST('testDeleteClearsTheCallersPointer');
	TraceStateFactory.parse(pDest:=pTraceState, pHeader:=ADR(traceState));
	THIS^._fillIds(traceId:=traceId, spanId:=spanId, seed:=0);
	ContextFactory.buildContext(
		pDest:=pContext,
		pTraceId:=ADR(traceId),
		pSpanId:=ADR(spanId),
		pTraceState:=pTraceState,
		traceFlags:=0
	);
	IF pTraceState <> 0 THEN pTraceState^.delete(pSelf:=pTraceState); END_IF
	IF pContext = 0 THEN
		THIS^.AssertTrue(FALSE, 'Expected buildContext to succeed');
		TcUnit.TEST_FINISHED();
		RETURN;
	END_IF

	deleted := pContext^.delete(pSelf:=pContext);
	THIS^.AssertTrue(deleted, 'Expected delete to report that the context was released');
	THIS^.AssertTrue(pContext = 0, 'Expected delete to clear the pointer of the caller');
TcUnit.TEST_FINISHED();
END_METHOD

(* delete only clears a pointer to the context it is called on. Handed a pointer to a different
   context, it must release nothing and leave both contexts and both pointers untouched. *)
METHOD testDeleteRefusesAnotherPointer : REFERENCE TO FB_Test
VAR
	pFirst: POINTER TO FB_SpanContext;
	pSecond: POINTER TO FB_SpanContext;
	pSecondBefore: POINTER TO FB_SpanContext;
	traceId: FB_TraceId;
	spanId: FB_SpanId;
	deleted: BOOL;
END_VAR
TcUnit.TEST('testDeleteRefusesAnotherPointer');
	THIS^._fillIds(traceId:=traceId, spanId:=spanId, seed:=0);
	ContextFactory.buildContext(pDest:=pFirst, pTraceId:=ADR(traceId), pSpanId:=ADR(spanId), pTraceState:=0, traceFlags:=0);
	ContextFactory.buildContext(pDest:=pSecond, pTraceId:=ADR(traceId), pSpanId:=ADR(spanId), pTraceState:=0, traceFlags:=0);
	IF pFirst = 0 OR pSecond = 0 THEN
		THIS^.AssertTrue(FALSE, 'Expected both builds to succeed');
		THIS^._release(pContext:=pFirst);
		THIS^._release(pContext:=pSecond);
		TcUnit.TEST_FINISHED();
		RETURN;
	END_IF
	pSecondBefore := pSecond;

	deleted := pFirst^.delete(pSelf:=pSecond);
	THIS^.AssertFalse(deleted, 'Expected delete to refuse a pointer to another context');
	THIS^.AssertTrue(pSecond = pSecondBefore, 'Expected the other pointer to be left untouched');
	THIS^.AssertTrue(pFirst^.isValid(), 'Expected the context not to be released');
	THIS^.AssertTrue(pSecond^.isValid(), 'Expected the other context not to be released');

	THIS^._release(pContext:=pFirst);
	THIS^._release(pContext:=pSecond);
TcUnit.TEST_FINISHED();
END_METHOD

(* free releases the trace state and clears the identity. Freeing twice must be harmless,
   and delete must still release a freed context. *)
METHOD testFreeClearsTheContext : REFERENCE TO FB_Test
VAR
	pContext: POINTER TO FB_SpanContext;
	traceId: FB_TraceId;
	spanId: FB_SpanId;
	traceState: T_MaxString := 'vendor=abc';
	pTraceState: POINTER TO FB_TraceState;
	success: BOOL;
END_VAR
TcUnit.TEST('testFreeClearsTheContext');
	TraceStateFactory.parse(pDest:=pTraceState, pHeader:=ADR(traceState));
	THIS^._fillIds(traceId:=traceId, spanId:=spanId, seed:=0);
	success := ContextFactory.buildContext(
		pDest:=pContext,
		pTraceId:=ADR(traceId),
		pSpanId:=ADR(spanId),
		pTraceState:=pTraceState,
		traceFlags:=16#301  // sampled, remoteness known, remote: every flag free must clear
	);
	IF pTraceState <> 0 THEN pTraceState^.delete(pSelf:=pTraceState); END_IF
	THIS^.AssertTrue(success, 'Expected buildContext to succeed');
	IF pContext = 0 THEN
		TcUnit.TEST_FINISHED();
		RETURN;
	END_IF

	pContext^.free();
	THIS^.AssertFalse(pContext^.isValid(), 'Expected a freed context to be invalid');
	THIS^.AssertFalse(pContext^.isRemote(), 'Expected a freed context not to report remote');
	THIS^.AssertTrue(pContext^.traceState = 0, 'Expected free to release the trace state');
	THIS^.AssertEquals_UDINT(0, pContext^.traceFlags, 'Expected free to clear the flags');

	pContext^.free();
	THIS^.AssertFalse(pContext^.isValid(), 'Expected a second free to leave the context empty');

	THIS^._release(pContext:=pContext);
	THIS^.AssertTrue(pContext = 0, 'Expected delete to clear the pointer');
TcUnit.TEST_FINISHED();
END_METHOD

(* Bit 8 says remoteness is known and bit 9 says the span is remote; only both together mean
   remote. The W3C trace flags in bits 0-7 must not affect the answer. *)
METHOD testIsRemoteNeedsBothBits : REFERENCE TO FB_Test
VAR
	pContext: POINTER TO FB_SpanContext;
	traceId: FB_TraceId;
	spanId: FB_SpanId;
	hasIsRemote: UDINT;
	isRemote: UDINT;
END_VAR
TcUnit.TEST('testIsRemoteNeedsBothBits');
	THIS^._fillIds(traceId:=traceId, spanId:=spanId, seed:=0);
	hasIsRemote := TO_UDINT(E_SpanFlags.SPAN_FLAGS_CONTEXT_HAS_IS_REMOTE_MASK);
	isRemote := TO_UDINT(E_SpanFlags.SPAN_FLAGS_CONTEXT_IS_REMOTE_MASK);

	ContextFactory.buildContext(pDest:=pContext, pTraceId:=ADR(traceId), pSpanId:=ADR(spanId), pTraceState:=0, traceFlags:=0);
	THIS^.AssertTrue(pContext <> 0 AND_THEN NOT pContext^.isRemote(), 'Expected no remoteness bits to mean not remote');
	THIS^._release(pContext:=pContext);

	ContextFactory.buildContext(pDest:=pContext, pTraceId:=ADR(traceId), pSpanId:=ADR(spanId), pTraceState:=0, traceFlags:=hasIsRemote);
	THIS^.AssertTrue(pContext <> 0 AND_THEN NOT pContext^.isRemote(), 'Expected known-and-local to mean not remote');
	THIS^._release(pContext:=pContext);

	ContextFactory.buildContext(pDest:=pContext, pTraceId:=ADR(traceId), pSpanId:=ADR(spanId), pTraceState:=0, traceFlags:=isRemote);
	THIS^.AssertTrue(pContext <> 0 AND_THEN NOT pContext^.isRemote(), 'Expected the remote bit without the known bit to mean not remote');
	THIS^._release(pContext:=pContext);

	ContextFactory.buildContext(pDest:=pContext, pTraceId:=ADR(traceId), pSpanId:=ADR(spanId), pTraceState:=0, traceFlags:=hasIsRemote OR isRemote);
	THIS^.AssertTrue(pContext <> 0 AND_THEN pContext^.isRemote(), 'Expected known-and-remote to mean remote');
	THIS^._release(pContext:=pContext);

	// 16#FF sets every W3C trace flag bit
	ContextFactory.buildContext(pDest:=pContext, pTraceId:=ADR(traceId), pSpanId:=ADR(spanId), pTraceState:=0, traceFlags:=hasIsRemote OR isRemote OR 16#FF);
	THIS^.AssertTrue(pContext <> 0 AND_THEN pContext^.isRemote(), 'Expected the W3C trace flags not to change the remote answer');
	THIS^._release(pContext:=pContext);
TcUnit.TEST_FINISHED();
END_METHOD

(* Like ValueFactory, buildContext never overwrites a pointer the caller already owns.
   A second build into the same destination must fail and leave the first context untouched. *)
METHOD testRejectsAssignedDestination : REFERENCE TO FB_Test
VAR
	pContext: POINTER TO FB_SpanContext;
	pFirst: POINTER TO FB_SpanContext;
	traceId: FB_TraceId;
	spanId: FB_SpanId;
	otherTraceId: FB_TraceId;
	otherSpanId: FB_SpanId;
	traceState: T_MaxString := 'vendor=abc';
	otherTraceState: T_MaxString := 'vendor=xyz';
	pTraceState: POINTER TO FB_TraceState;
	pOtherTraceState: POINTER TO FB_TraceState;
	success: BOOL;
	failureReason: E_ContextFactoryFailureReason;
END_VAR
TcUnit.TEST('testRejectsAssignedDestination');
	TraceStateFactory.parse(pDest:=pTraceState, pHeader:=ADR(traceState));
	TraceStateFactory.parse(pDest:=pOtherTraceState, pHeader:=ADR(otherTraceState));
	THIS^._fillIds(traceId:=traceId, spanId:=spanId, seed:=0);
	THIS^._fillIds(traceId:=otherTraceId, spanId:=otherSpanId, seed:=16#80);

	success := ContextFactory.buildContext(
		pDest:=pContext,
		pTraceId:=ADR(traceId),
		pSpanId:=ADR(spanId),
		pTraceState:=pTraceState,
		traceFlags:=1  // sampled, so the kept flags can be told from the second build's 0
	);
	IF pTraceState <> 0 THEN pTraceState^.delete(pSelf:=pTraceState); END_IF
	THIS^.AssertTrue(success, 'Expected the first build to succeed');
	IF pContext = 0 THEN
		IF pOtherTraceState <> 0 THEN pOtherTraceState^.delete(pSelf:=pOtherTraceState); END_IF
		TcUnit.TEST_FINISHED();
		RETURN;
	END_IF
	pFirst := pContext;

	success := ContextFactory.buildContext(
		pDest:=pContext,
		pTraceId:=ADR(otherTraceId),
		pSpanId:=ADR(otherSpanId),
		pTraceState:=pOtherTraceState,
		traceFlags:=0,
		failureReason=>failureReason
	);
	IF pOtherTraceState <> 0 THEN pOtherTraceState^.delete(pSelf:=pOtherTraceState); END_IF
	THIS^.AssertFalse(success, 'Expected a build into an assigned destination to fail');
	THIS^.AssertEquals_UDINT(
		TO_UDINT(E_ContextFactoryFailureReason.DESTINATION_ALREADY_ASSIGNED),
		TO_UDINT(failureReason),
		'Expected an assigned destination to report DESTINATION_ALREADY_ASSIGNED'
	);
	THIS^.AssertTrue(pContext = pFirst, 'Expected the destination pointer to be left alone');
	THIS^.AssertTrue(
		MEMCMP(ADR(pContext^.spanId.bytes), ADR(spanId.bytes), SIZEOF(spanId.bytes)) = 0,
		'Expected the original span id to be kept'
	);
	THIS^.AssertEquals_UDINT(1, pContext^.traceFlags, 'Expected the original flags to be kept');
	IF pContext^.traceState <> 0 THEN
		THIS^.AssertEquals_STRING('vendor=abc', pContext^.traceState^.pString^, 'Expected the original trace state to be kept');
	ELSE
		THIS^.AssertTrue(FALSE, 'Expected the original trace state to be kept');
	END_IF

	THIS^._release(pContext:=pContext);
TcUnit.TEST_FINISHED();
END_METHOD

(* A null identifier pointer is a caller error, not an invalid identity. buildContext must
   refuse it without allocating anything. *)
METHOD testRejectsNullIdentifiers : REFERENCE TO FB_Test
VAR
	pContext: POINTER TO FB_SpanContext;
	traceId: FB_TraceId;
	spanId: FB_SpanId;
	traceState: T_MaxString := 'vendor=abc';
	pTraceState: POINTER TO FB_TraceState;
	success: BOOL;
	failureReason: E_ContextFactoryFailureReason;
END_VAR
TcUnit.TEST('testRejectsNullIdentifiers');
	TraceStateFactory.parse(pDest:=pTraceState, pHeader:=ADR(traceState));
	THIS^._fillIds(traceId:=traceId, spanId:=spanId, seed:=0);

	success := ContextFactory.buildContext(
		pDest:=pContext,
		pTraceId:=0,
		pSpanId:=ADR(spanId),
		pTraceState:=pTraceState,
		traceFlags:=1,
		failureReason=>failureReason
	);
	THIS^.AssertFalse(success, 'Expected buildContext to reject a null trace id pointer');
	THIS^.AssertEquals_UDINT(
		TO_UDINT(E_ContextFactoryFailureReason.TRACE_ID_POINTER_NULL),
		TO_UDINT(failureReason),
		'Expected a null trace id pointer to report TRACE_ID_POINTER_NULL'
	);
	THIS^.AssertTrue(pContext = 0, 'Expected a rejected build to leave the destination unassigned');

	success := ContextFactory.buildContext(
		pDest:=pContext,
		pTraceId:=ADR(traceId),
		pSpanId:=0,
		pTraceState:=pTraceState,
		traceFlags:=1,
		failureReason=>failureReason
	);
	THIS^.AssertFalse(success, 'Expected buildContext to reject a null span id pointer');
	THIS^.AssertEquals_UDINT(
		TO_UDINT(E_ContextFactoryFailureReason.SPAN_ID_POINTER_NULL),
		TO_UDINT(failureReason),
		'Expected a null span id pointer to report SPAN_ID_POINTER_NULL'
	);
	THIS^.AssertTrue(pContext = 0, 'Expected a rejected build to leave the destination unassigned');

	IF pTraceState <> 0 THEN pTraceState^.delete(pSelf:=pTraceState); END_IF
	THIS^._release(pContext:=pContext);
TcUnit.TEST_FINISHED();
END_METHOD

(* fromSpan refuses a null span without allocating anything. *)
METHOD testFromSpanRejectsNullSpan : REFERENCE TO FB_Test
VAR
	pContext: POINTER TO FB_SpanContext;
	success: BOOL;
	failureReason: E_ContextFactoryFailureReason;
END_VAR
TcUnit.TEST('testFromSpanRejectsNullSpan');
	success := ContextFactory.fromSpan(pDest:=pContext, pSpan:=0, failureReason=>failureReason);
	THIS^.AssertFalse(success, 'Expected fromSpan to refuse a null span');
	THIS^.AssertEquals_UDINT(
		TO_UDINT(E_ContextFactoryFailureReason.SPAN_POINTER_NULL),
		TO_UDINT(failureReason),
		'Expected SPAN_POINTER_NULL'
	);
	THIS^.AssertTrue(pContext = 0, 'Expected the destination to stay unassigned');
TcUnit.TEST_FINISHED();
END_METHOD

END_FUNCTION_BLOCK

// ---- TEST/TRACING/TRACESTATE/FB_TestTraceState.TcPOU
(* Tests TraceStateFactory and FB_TraceState against the W3C tracestate rules. *)
FUNCTION_BLOCK FB_TestTraceState EXTENDS FB_TestSuite

THIS^.testParseCanonicalises();
THIS^.testParseEmptyHeader();
THIS^.testParseRejectsInvalidHeaders();
THIS^.testParseEntryLimit();
THIS^.testParseLongHeader();
THIS^.testCloneIsIndependent();
THIS^.testTruncateFollowsW3C();

